// LS Electric XG5000 project: eduPJT_A
// PLC LSPLC
// module base 0 slot 0: 입출력 모듈:XBC-DR32H (DC 24V 입력, 릴레이 출력 32점)
// module base 0 slot 1: 입력 모듈:XBE-DC16A/B (DC24V 입력, 16점 / DC12/24V 입력, 16점)
// module base 0 slot 2: FEnet:XBL-EMTA (Ethernet 통신 모듈, 전기 Master)

PROGRAM 00_Global_Layer (task: 스캔 프로그램)

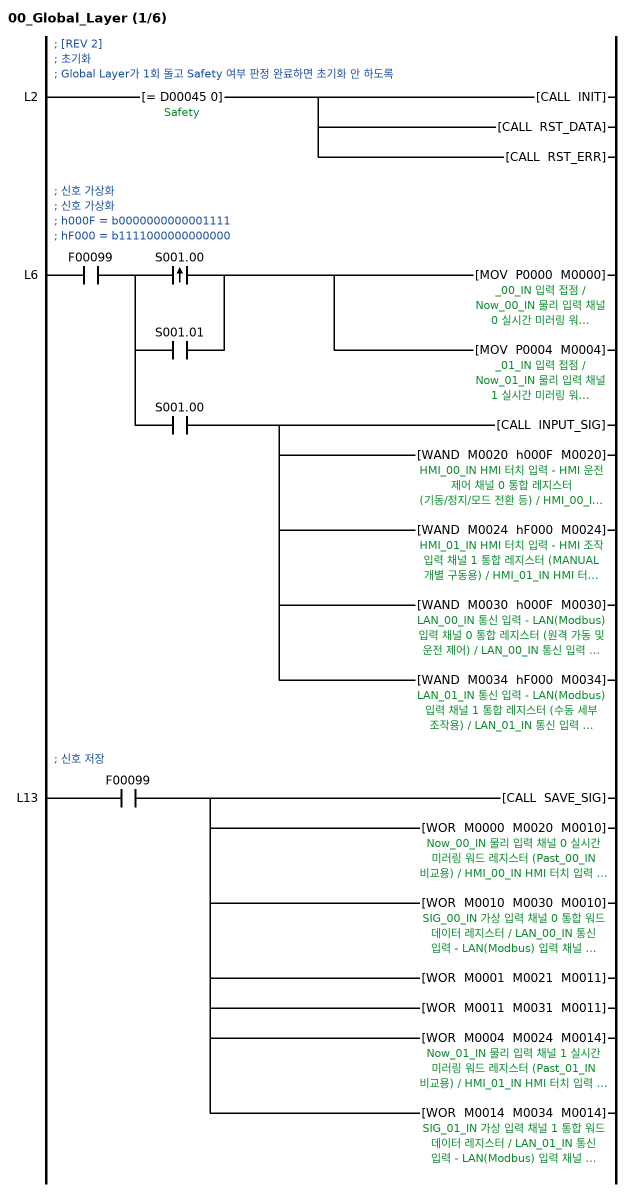
// [REV 2]
// 초기화
; L2
LOAD=     D00045 0	// Safety
CALL      INIT
CALL      RST_DATA
CALL      RST_ERR
// output comment: Global Layer가 1회 돌고 Safety 여부 판정 완료하면 초기화 안 하도록
// 신호 가상화
; L6
LOAD      F00099
MPUSH
LOADP     S001.00
OR        S001.01
AND LOAD
MOV       P0000 M0000	// _00_IN 입력 접점 / Now_00_IN 물리 입력 채널 0 실시간 미러링 워드 레지스터 (Past_00_IN 비교용)
MOV       P0004 M0004	// _01_IN 입력 접점 / Now_01_IN 물리 입력 채널 1 실시간 미러링 워드 레지스터 (Past_01_IN 비교용)
MPOP
AND       S001.00
CALL      INPUT_SIG
WAND      M0020 h000F M0020	// HMI_00_IN HMI 터치 입력 - HMI 운전 제어 채널 0 통합 레지스터 (기동/정지/모드 전환 등) / HMI_00_IN HMI 터치 입력 - HMI 운전 제어 채널 0 통합 레지스터 (기동/정지/모드 전환 등)
WAND      M0024 hF000 M0024	// HMI_01_IN HMI 터치 입력 - HMI 조작 입력 채널 1 통합 레지스터 (MANUAL 개별 구동용) / HMI_01_IN HMI 터치 입력 - HMI 조작 입력 채널 1 통합 레지스터 (MANUAL 개별 구동용)
WAND      M0030 h000F M0030	// LAN_00_IN 통신 입력 - LAN(Modbus) 입력 채널 0 통합 레지스터 (원격 가동 및 운전 제어) / LAN_00_IN 통신 입력 - LAN(Modbus) 입력 채널 0 통합 레지스터 (원격 가동 및 운전 제어)
WAND      M0034 hF000 M0034	// LAN_01_IN 통신 입력 - LAN(Modbus) 입력 채널 1 통합 레지스터 (수동 세부 조작용) / LAN_01_IN 통신 입력 - LAN(Modbus) 입력 채널 1 통합 레지스터 (수동 세부 조작용)
// output comment: 신호 가상화
// output comment: h000F = b0000000000001111
// output comment: hF000 = b1111000000000000
; L13
LOAD      F00099
CALL      SAVE_SIG
WOR       M0000 M0020 M0010	// Now_00_IN 물리 입력 채널 0 실시간 미러링 워드 레지스터 (Past_00_IN 비교용) / HMI_00_IN HMI 터치 입력 - HMI 운전 제어 채널 0 통합 레지스터 (기동/정지/모드 전환 등) / SIG_00_IN 가상 입력 채널 0 통합 워드 데이터 레지스터
WOR       M0010 M0030 M0010	// SIG_00_IN 가상 입력 채널 0 통합 워드 데이터 레지스터 / LAN_00_IN 통신 입력 - LAN(Modbus) 입력 채널 0 통합 레지스터 (원격 가동 및 운전 제어) / SIG_00_IN 가상 입력 채널 0 통합 워드 데이터 레지스터
WOR       M0001 M0021 M0011
WOR       M0011 M0031 M0011
WOR       M0004 M0024 M0014	// Now_01_IN 물리 입력 채널 1 실시간 미러링 워드 레지스터 (Past_01_IN 비교용) / HMI_01_IN HMI 터치 입력 - HMI 조작 입력 채널 1 통합 레지스터 (MANUAL 개별 구동용) / SIG_01_IN 가상 입력 채널 1 통합 워드 데이터 레지스터
WOR       M0014 M0034 M0014	// SIG_01_IN 가상 입력 채널 1 통합 워드 데이터 레지스터 / LAN_01_IN 통신 입력 - LAN(Modbus) 입력 채널 1 통합 레지스터 (수동 세부 조작용) / SIG_01_IN 가상 입력 채널 1 통합 워드 데이터 레지스터
// output comment: 신호 저장

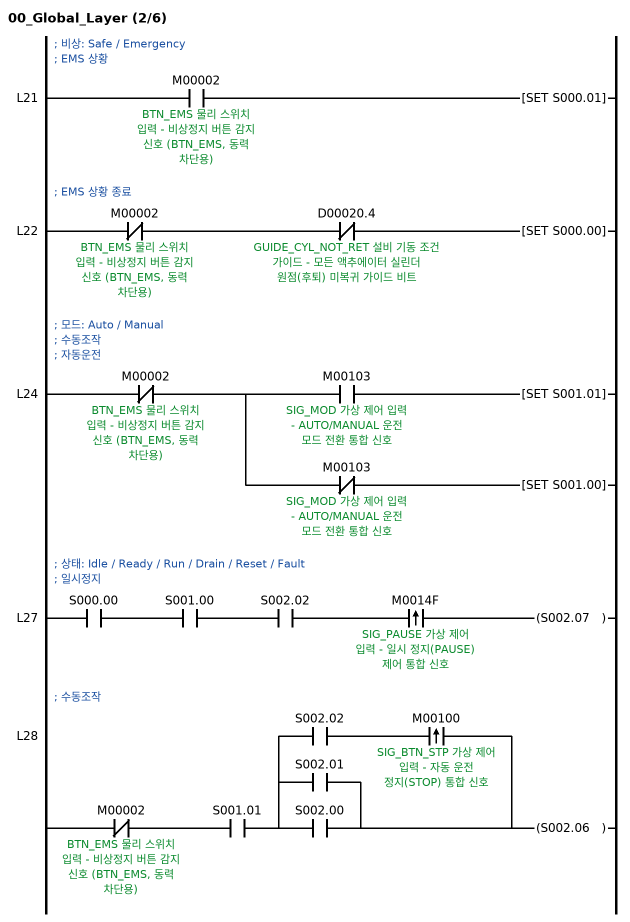
// 비상: Safe / Emergency
; L21
LOAD      M00002	// BTN_EMS 물리 스위치 입력 - 비상정지 버튼 감지 신호 (BTN_EMS, 동력 차단용)
SET       S000.01
// output comment: EMS 상황
; L22
LOAD NOT  M00002	// BTN_EMS 물리 스위치 입력 - 비상정지 버튼 감지 신호 (BTN_EMS, 동력 차단용)
AND NOT   D00020.4	// GUIDE_CYL_NOT_RET 설비 기동 조건 가이드 - 모든 액추에이터 실린더 원점(후퇴) 미복귀 가이드 비트
SET       S000.00
// output comment: EMS 상황 종료
// 모드: Auto / Manual
; L24
LOAD NOT  M00002	// BTN_EMS 물리 스위치 입력 - 비상정지 버튼 감지 신호 (BTN_EMS, 동력 차단용)
MPUSH
AND       M00103	// SIG_MOD 가상 제어 입력 - AUTO/MANUAL 운전 모드 전환 통합 신호
SET       S001.01
MPOP
AND NOT   M00103	// SIG_MOD 가상 제어 입력 - AUTO/MANUAL 운전 모드 전환 통합 신호
SET       S001.00
// output comment: 수동조작
// output comment: 자동운전
// 상태: Idle / Ready / Run / Drain / Reset / Fault
; L27
LOAD      S000.00
AND       S001.00
AND       S002.02
ANDP      M0014F	// SIG_PAUSE 가상 제어 입력 - 일시 정지(PAUSE) 제어 통합 신호
OUT       S002.07
// output comment: 일시정지
; L28
LOAD NOT  M00002	// BTN_EMS 물리 스위치 입력 - 비상정지 버튼 감지 신호 (BTN_EMS, 동력 차단용)
AND       S001.01
LOAD      S002.02
ANDP      M00100	// SIG_BTN_STP 가상 제어 입력 - 자동 운전 정지(STOP) 통합 신호
OR        S002.01
OR        S002.00
AND LOAD
OUT       S002.06
// output comment: 수동조작

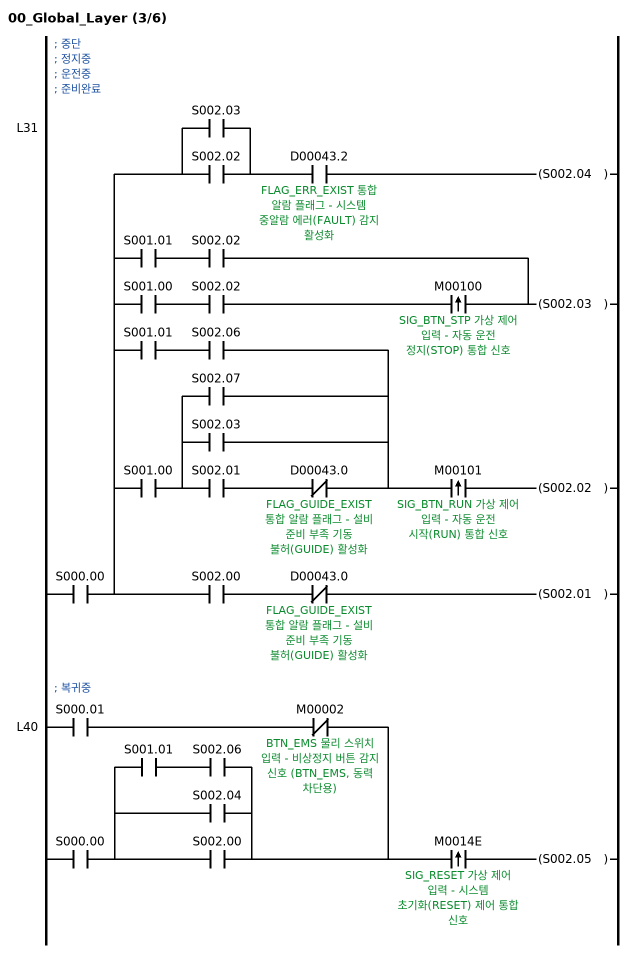
; L31
LOAD      S000.00
MPUSH
LOAD      S002.03
OR        S002.02
AND LOAD
AND       D00043.2	// FLAG_ERR_EXIST 통합 알람 플래그 - 시스템 중알람 에러(FAULT) 감지 활성화
OUT       S002.04
MLOAD
LOAD      S001.01
AND       S002.02
LOAD      S001.00
AND       S002.02
ANDP      M00100	// SIG_BTN_STP 가상 제어 입력 - 자동 운전 정지(STOP) 통합 신호
OR LOAD
AND LOAD
OUT       S002.03
MLOAD
LOAD      S001.01
AND       S002.06
LOAD      S001.00
LOAD      S002.07
OR        S002.03
LOAD      S002.01
AND NOT   D00043.0	// FLAG_GUIDE_EXIST 통합 알람 플래그 - 설비 준비 부족 기동 불허(GUIDE) 활성화
OR LOAD
AND LOAD
OR LOAD
AND LOAD
ANDP      M00101	// SIG_BTN_RUN 가상 제어 입력 - 자동 운전 시작(RUN) 통합 신호
OUT       S002.02
MPOP
AND       S002.00
AND NOT   D00043.0	// FLAG_GUIDE_EXIST 통합 알람 플래그 - 설비 준비 부족 기동 불허(GUIDE) 활성화
OUT       S002.01
// output comment: 중단
// output comment: 정지중
// output comment: 운전중
// output comment: 준비완료
; L40
LOAD      S000.01
AND NOT   M00002	// BTN_EMS 물리 스위치 입력 - 비상정지 버튼 감지 신호 (BTN_EMS, 동력 차단용)
LOAD      S000.00
LOAD      S001.01
AND       S002.06
OR        S002.04
OR        S002.00
AND LOAD
OR LOAD
ANDP      M0014E	// SIG_RESET 가상 제어 입력 - 시스템 초기화(RESET) 제어 통합 신호
OUT       S002.05
// output comment: 복귀중

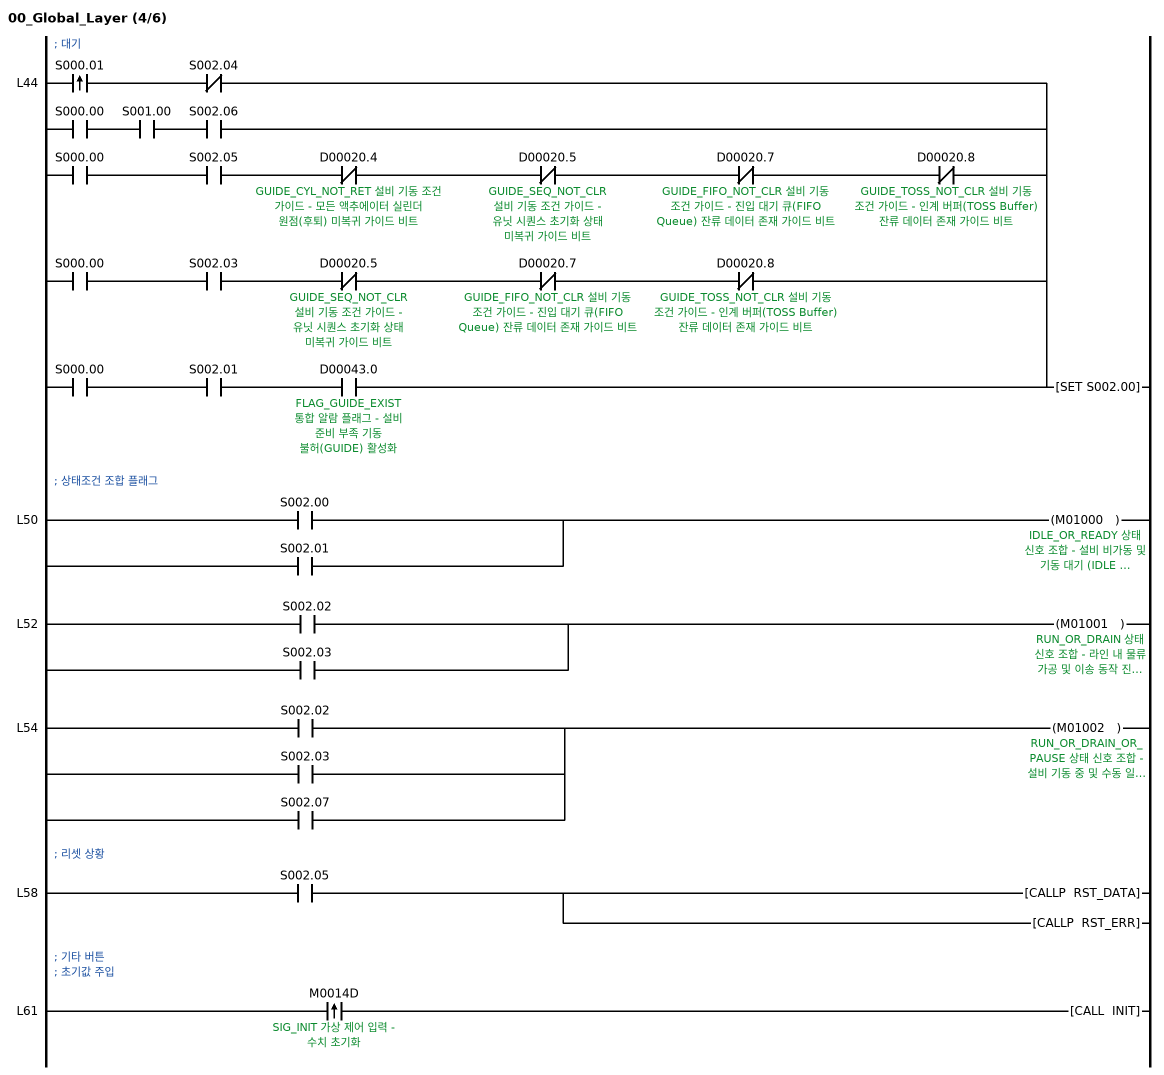
; L44
LOADP     S000.01
AND NOT   S002.04
LOAD      S000.00
AND       S001.00
AND       S002.06
OR LOAD
LOAD      S000.00
AND       S002.05
AND NOT   D00020.4	// GUIDE_CYL_NOT_RET 설비 기동 조건 가이드 - 모든 액추에이터 실린더 원점(후퇴) 미복귀 가이드 비트
AND NOT   D00020.5	// GUIDE_SEQ_NOT_CLR 설비 기동 조건 가이드 - 유닛 시퀀스 초기화 상태 미복귀 가이드 비트
AND NOT   D00020.7	// GUIDE_FIFO_NOT_CLR 설비 기동 조건 가이드 - 진입 대기 큐(FIFO Queue) 잔류 데이터 존재 가이드 비트
AND NOT   D00020.8	// GUIDE_TOSS_NOT_CLR 설비 기동 조건 가이드 - 인계 버퍼(TOSS Buffer) 잔류 데이터 존재 가이드 비트
OR LOAD
LOAD      S000.00
AND       S002.03
AND NOT   D00020.5	// GUIDE_SEQ_NOT_CLR 설비 기동 조건 가이드 - 유닛 시퀀스 초기화 상태 미복귀 가이드 비트
AND NOT   D00020.7	// GUIDE_FIFO_NOT_CLR 설비 기동 조건 가이드 - 진입 대기 큐(FIFO Queue) 잔류 데이터 존재 가이드 비트
AND NOT   D00020.8	// GUIDE_TOSS_NOT_CLR 설비 기동 조건 가이드 - 인계 버퍼(TOSS Buffer) 잔류 데이터 존재 가이드 비트
OR LOAD
LOAD      S000.00
AND       S002.01
AND       D00043.0	// FLAG_GUIDE_EXIST 통합 알람 플래그 - 설비 준비 부족 기동 불허(GUIDE) 활성화
OR LOAD
SET       S002.00
// output comment: 대기
// 상태조건 조합 플래그
; L50
LOAD      S002.00
OR        S002.01
OUT       M01000	// IDLE_OR_READY 상태 신호 조합 - 설비 비가동 및 기동 대기 (IDLE | READY) 플래그
; L52
LOAD      S002.02
OR        S002.03
OUT       M01001	// RUN_OR_DRAIN 상태 신호 조합 - 라인 내 물류 가공 및 이송 동작 진행 (RUN | DRAIN) 플래그
; L54
LOAD      S002.02
OR        S002.03
OR        S002.07
OUT       M01002	// RUN_OR_DRAIN_OR_PAUSE 상태 신호 조합 - 설비 기동 중 및 수동 일시 정지 (RUN | DRAIN | PAUSE) 플래그
// 리셋 상황
; L58
LOAD      S002.05
CALLP     RST_DATA
CALLP     RST_ERR
// 기타 버튼
; L61
LOADP     M0014D	// SIG_INIT 가상 제어 입력 - 수치 초기화
CALL      INIT
// output comment: 초기값 주입

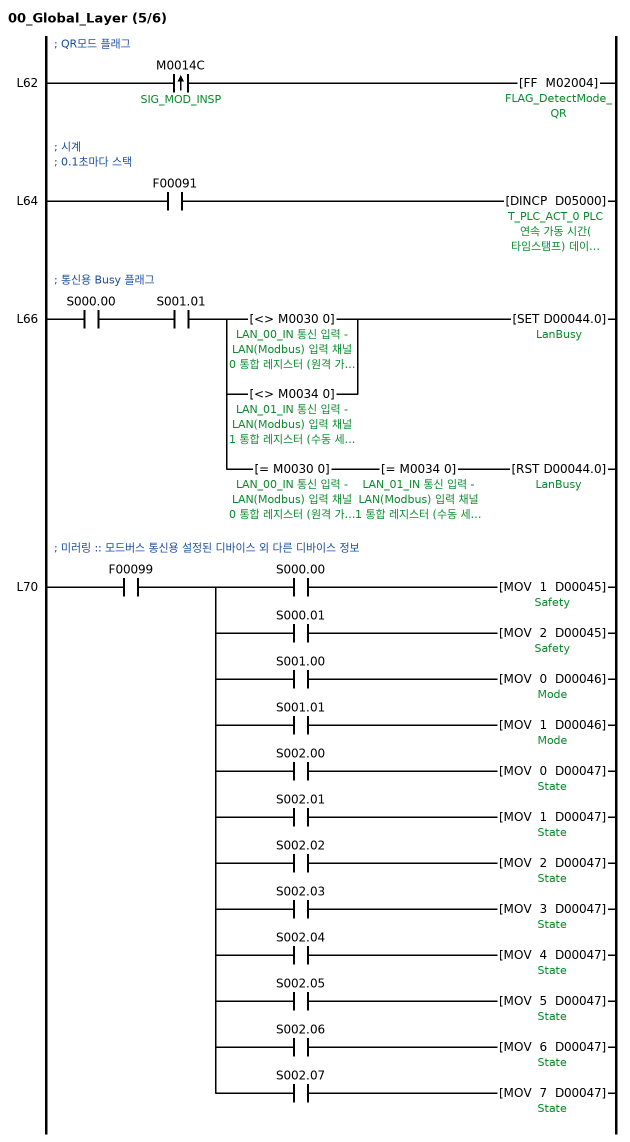
; L62
LOADP     M0014C	// SIG_MOD_INSP
FF        M02004	// FLAG_DetectMode_QR
// output comment: QR모드 플래그
// 시계
; L64
LOAD      F00091
DINCP     D05000	// T_PLC_ACT_0 PLC 연속 가동 시간(타임스탬프) 데이터 레지스터 하위 16비트 (0.1초 해상도)
// output comment: 0.1초마다 스택
// 통신용 Busy 플래그
; L66
LOAD      S000.00
AND       S001.01
MPUSH
LOAD<>    M0030 0	// LAN_00_IN 통신 입력 - LAN(Modbus) 입력 채널 0 통합 레지스터 (원격 가동 및 운전 제어)
OR<>      M0034 0	// LAN_01_IN 통신 입력 - LAN(Modbus) 입력 채널 1 통합 레지스터 (수동 세부 조작용)
AND LOAD
SET       D00044.0	// LanBusy
MPOP
AND=      M0030 0	// LAN_00_IN 통신 입력 - LAN(Modbus) 입력 채널 0 통합 레지스터 (원격 가동 및 운전 제어)
AND=      M0034 0	// LAN_01_IN 통신 입력 - LAN(Modbus) 입력 채널 1 통합 레지스터 (수동 세부 조작용)
RST       D00044.0	// LanBusy
// 미러링 :: 모드버스 통신용 설정된 디바이스 외 다른 디바이스 정보
; L70
LOAD      F00099
MPUSH
AND       S000.00
MOV       1 D00045	// Safety
MLOAD
AND       S000.01
MOV       2 D00045	// Safety
MLOAD
AND       S001.00
MOV       0 D00046	// Mode
MLOAD
AND       S001.01
MOV       1 D00046	// Mode
MLOAD
AND       S002.00
MOV       0 D00047	// State
MLOAD
AND       S002.01
MOV       1 D00047	// State
MLOAD
AND       S002.02
MOV       2 D00047	// State
MLOAD
AND       S002.03
MOV       3 D00047	// State
MLOAD
AND       S002.04
MOV       4 D00047	// State
MLOAD
AND       S002.05
MOV       5 D00047	// State
MLOAD
AND       S002.06
MOV       6 D00047	// State
MPOP
AND       S002.07
MOV       7 D00047	// State

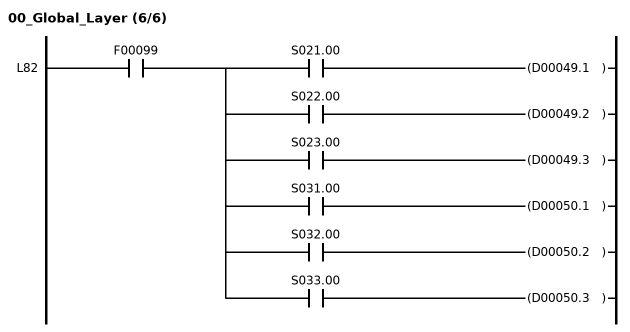
; L82
LOAD      F00099
MPUSH
AND       S021.00
OUT       D00049.1
MLOAD
AND       S022.00
OUT       D00049.2
MLOAD
AND       S023.00
OUT       D00049.3
MLOAD
AND       S031.00
OUT       D00050.1
MLOAD
AND       S032.00
OUT       D00050.2
MPOP
AND       S033.00
OUT       D00050.3

PROGRAM 01_Sequence_Layer (task: 스캔 프로그램)

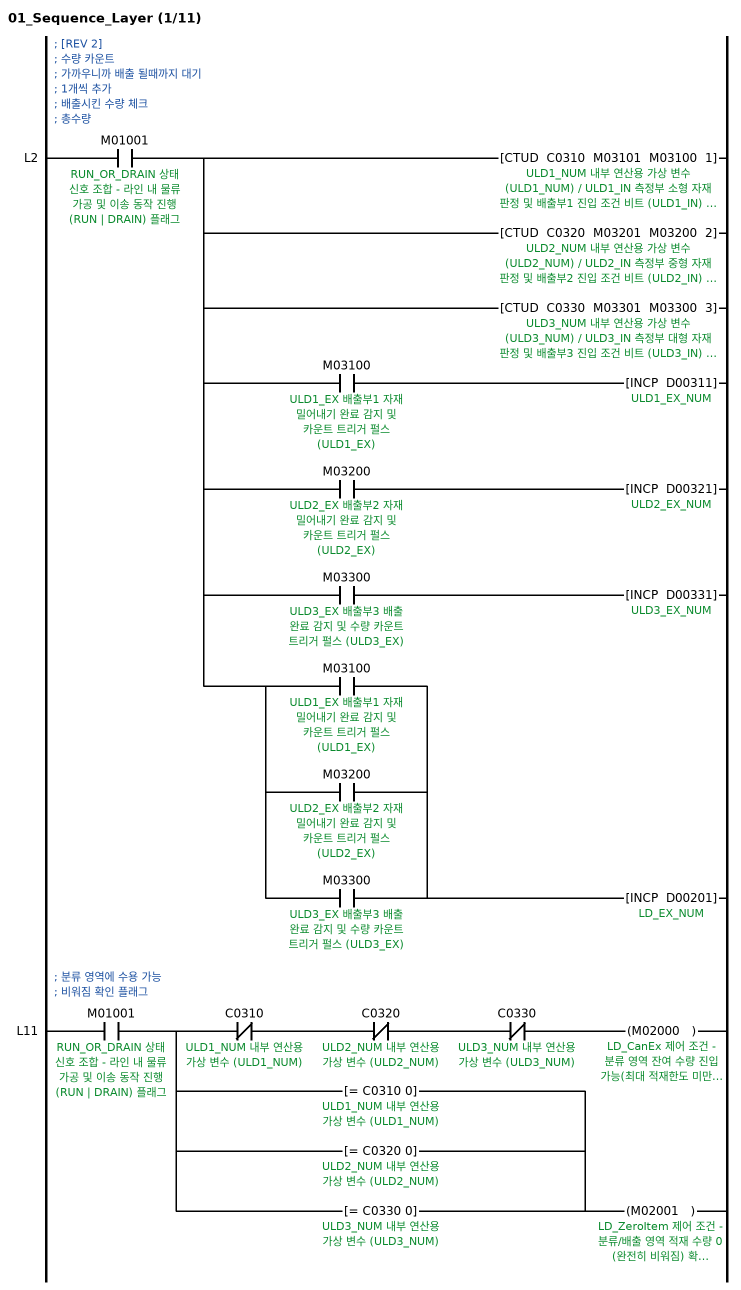
// [REV 2]
// 수량 카운트
; L2
LOAD      M01001	// RUN_OR_DRAIN 상태 신호 조합 - 라인 내 물류 가공 및 이송 동작 진행 (RUN | DRAIN) 플래그
CTUD      C0310 M03101 M03100 1	// ULD1_NUM 내부 연산용 가상 변수 (ULD1_NUM) / ULD1_IN 측정부 소형 자재 판정 및 배출부1 진입 조건 비트 (ULD1_IN) / ULD1_EX 배출부1 자재 밀어내기 완료 감지 및 카운트 트리거 펄스 (ULD1_EX)
CTUD      C0320 M03201 M03200 2	// ULD2_NUM 내부 연산용 가상 변수 (ULD2_NUM) / ULD2_IN 측정부 중형 자재 판정 및 배출부2 진입 조건 비트 (ULD2_IN) / ULD2_EX 배출부2 자재 밀어내기 완료 감지 및 카운트 트리거 펄스 (ULD2_EX)
CTUD      C0330 M03301 M03300 3	// ULD3_NUM 내부 연산용 가상 변수 (ULD3_NUM) / ULD3_IN 측정부 대형 자재 판정 및 배출부3 진입 조건 비트 (ULD3_IN) / ULD3_EX 배출부3 배출 완료 감지 및 수량 카운트 트리거 펄스 (ULD3_EX)
MPUSH
AND       M03100	// ULD1_EX 배출부1 자재 밀어내기 완료 감지 및 카운트 트리거 펄스 (ULD1_EX)
INCP      D00311	// ULD1_EX_NUM
MLOAD
AND       M03200	// ULD2_EX 배출부2 자재 밀어내기 완료 감지 및 카운트 트리거 펄스 (ULD2_EX)
INCP      D00321	// ULD2_EX_NUM
MLOAD
AND       M03300	// ULD3_EX 배출부3 배출 완료 감지 및 수량 카운트 트리거 펄스 (ULD3_EX)
INCP      D00331	// ULD3_EX_NUM
MPOP
LOAD      M03100	// ULD1_EX 배출부1 자재 밀어내기 완료 감지 및 카운트 트리거 펄스 (ULD1_EX)
OR        M03200	// ULD2_EX 배출부2 자재 밀어내기 완료 감지 및 카운트 트리거 펄스 (ULD2_EX)
OR        M03300	// ULD3_EX 배출부3 배출 완료 감지 및 수량 카운트 트리거 펄스 (ULD3_EX)
AND LOAD
INCP      D00201	// LD_EX_NUM
// output comment: 가까우니까 배출 될때까지 대기
// output comment: 1개씩 추가
// output comment: 배출시킨 수량 체크
// output comment: 총수량
; L11
LOAD      M01001	// RUN_OR_DRAIN 상태 신호 조합 - 라인 내 물류 가공 및 이송 동작 진행 (RUN | DRAIN) 플래그
MPUSH
AND NOT   C0310	// ULD1_NUM 내부 연산용 가상 변수 (ULD1_NUM)
AND NOT   C0320	// ULD2_NUM 내부 연산용 가상 변수 (ULD2_NUM)
AND NOT   C0330	// ULD3_NUM 내부 연산용 가상 변수 (ULD3_NUM)
OUT       M02000	// LD_CanEx 제어 조건 - 분류 영역 잔여 수량 진입 가능(최대 적재한도 미만) 확인 플래그 (LD_CanEx)
MPOP
LOAD=     C0310 0	// ULD1_NUM 내부 연산용 가상 변수 (ULD1_NUM)
OR=       C0320 0	// ULD2_NUM 내부 연산용 가상 변수 (ULD2_NUM)
OR=       C0330 0	// ULD3_NUM 내부 연산용 가상 변수 (ULD3_NUM)
AND LOAD
OUT       M02001	// LD_ZeroItem 제어 조건 - 분류/배출 영역 적재 수량 0 (완전히 비워짐) 확인 플래그 (LD_ZeroItem)
// output comment: 분류 영역에 수용 가능
// output comment: 비워짐 확인 플래그

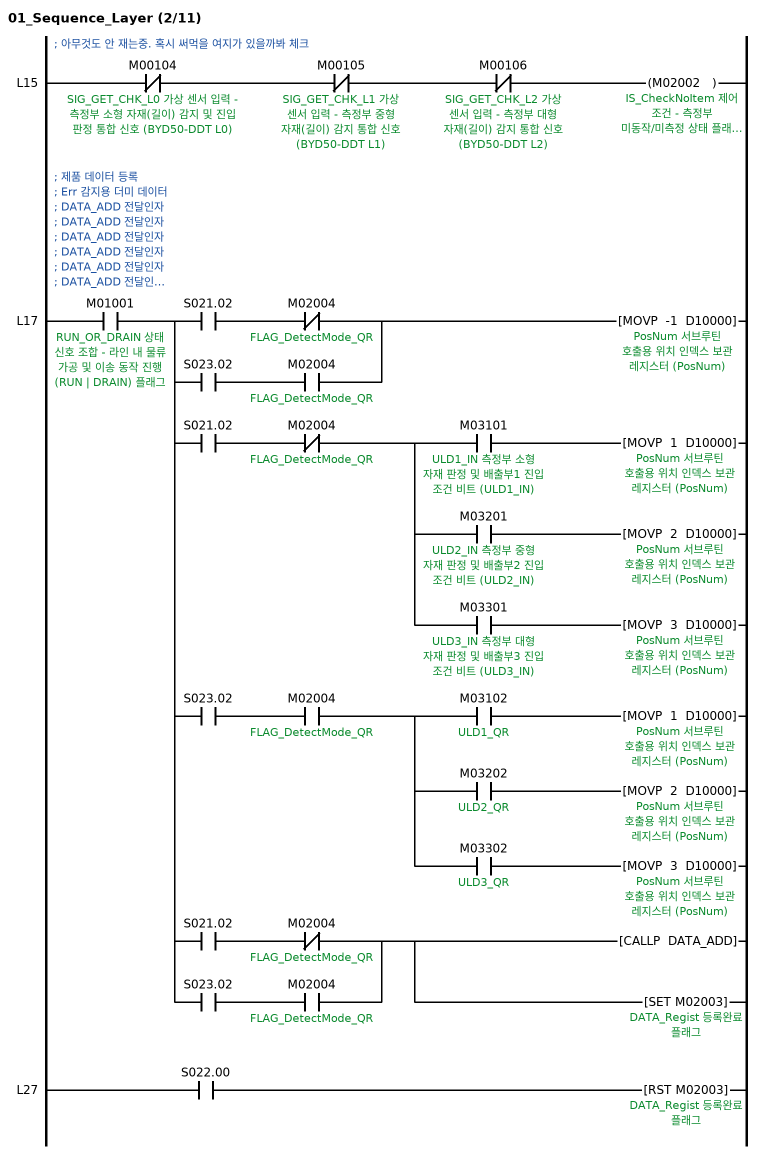
; L15
LOAD NOT  M00104	// SIG_GET_CHK_L0 가상 센서 입력 - 측정부 소형 자재(길이) 감지 및 진입 판정 통합 신호 (BYD50-DDT L0)
AND NOT   M00105	// SIG_GET_CHK_L1 가상 센서 입력 - 측정부 중형 자재(길이) 감지 통합 신호 (BYD50-DDT L1)
AND NOT   M00106	// SIG_GET_CHK_L2 가상 센서 입력 - 측정부 대형 자재(길이) 감지 통합 신호 (BYD50-DDT L2)
OUT       M02002	// IS_CheckNoItem 제어 조건 - 측정부 미동작/미측정 상태 플래그 (IS_CheckNoItem)
// output comment: 아무것도 안 재는중. 혹시 써먹을 여지가 있을까봐 체크
// 제품 데이터 등록
; L17
LOAD      M01001	// RUN_OR_DRAIN 상태 신호 조합 - 라인 내 물류 가공 및 이송 동작 진행 (RUN | DRAIN) 플래그
MPUSH
LOAD      S021.02
AND NOT   M02004	// FLAG_DetectMode_QR
LOAD      S023.02
AND       M02004	// FLAG_DetectMode_QR
OR LOAD
AND LOAD
MOVP      -1 D10000	// PosNum 서브루틴 호출용 위치 인덱스 보관 레지스터 (PosNum)
MLOAD
AND       S021.02
AND NOT   M02004	// FLAG_DetectMode_QR
MPUSH
AND       M03101	// ULD1_IN 측정부 소형 자재 판정 및 배출부1 진입 조건 비트 (ULD1_IN)
MOVP      1 D10000	// PosNum 서브루틴 호출용 위치 인덱스 보관 레지스터 (PosNum)
MLOAD
AND       M03201	// ULD2_IN 측정부 중형 자재 판정 및 배출부2 진입 조건 비트 (ULD2_IN)
MOVP      2 D10000	// PosNum 서브루틴 호출용 위치 인덱스 보관 레지스터 (PosNum)
MPOP
AND       M03301	// ULD3_IN 측정부 대형 자재 판정 및 배출부3 진입 조건 비트 (ULD3_IN)
MOVP      3 D10000	// PosNum 서브루틴 호출용 위치 인덱스 보관 레지스터 (PosNum)
MLOAD
AND       S023.02
AND       M02004	// FLAG_DetectMode_QR
MPUSH
AND       M03102	// ULD1_QR
MOVP      1 D10000	// PosNum 서브루틴 호출용 위치 인덱스 보관 레지스터 (PosNum)
MLOAD
AND       M03202	// ULD2_QR
MOVP      2 D10000	// PosNum 서브루틴 호출용 위치 인덱스 보관 레지스터 (PosNum)
MPOP
AND       M03302	// ULD3_QR
MOVP      3 D10000	// PosNum 서브루틴 호출용 위치 인덱스 보관 레지스터 (PosNum)
MPOP
LOAD      S021.02
AND NOT   M02004	// FLAG_DetectMode_QR
LOAD      S023.02
AND       M02004	// FLAG_DetectMode_QR
OR LOAD
AND LOAD
CALLP     DATA_ADD
SET       M02003	// DATA_Regist 등록완료 플래그
// output comment: Err 감지용 더미 데이터
// output comment: DATA_ADD 전달인자
// output comment: DATA_ADD 전달인자
// output comment: DATA_ADD 전달인자
// output comment: DATA_ADD 전달인자
// output comment: DATA_ADD 전달인자
// output comment: DATA_ADD 전달인자
// output comment: 선입선출 데이터 입력
// output comment: 등록완료 플래그
; L27
LOAD      S022.00
RST       M02003	// DATA_Regist 등록완료 플래그

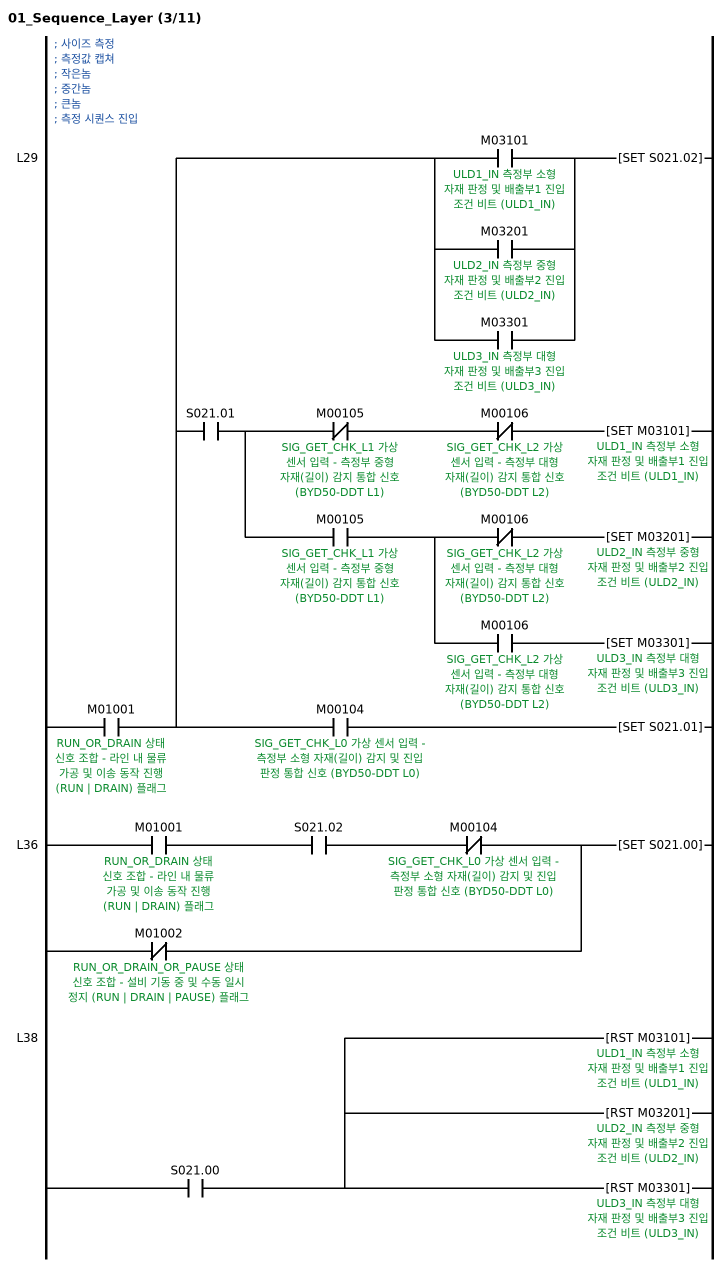
// 
// 사이즈 측정
; L29
LOAD      M01001	// RUN_OR_DRAIN 상태 신호 조합 - 라인 내 물류 가공 및 이송 동작 진행 (RUN | DRAIN) 플래그
MPUSH
LOAD      M03101	// ULD1_IN 측정부 소형 자재 판정 및 배출부1 진입 조건 비트 (ULD1_IN)
OR        M03201	// ULD2_IN 측정부 중형 자재 판정 및 배출부2 진입 조건 비트 (ULD2_IN)
OR        M03301	// ULD3_IN 측정부 대형 자재 판정 및 배출부3 진입 조건 비트 (ULD3_IN)
AND LOAD
SET       S021.02
MLOAD
AND       S021.01
MPUSH
AND NOT   M00105	// SIG_GET_CHK_L1 가상 센서 입력 - 측정부 중형 자재(길이) 감지 통합 신호 (BYD50-DDT L1)
AND NOT   M00106	// SIG_GET_CHK_L2 가상 센서 입력 - 측정부 대형 자재(길이) 감지 통합 신호 (BYD50-DDT L2)
SET       M03101	// ULD1_IN 측정부 소형 자재 판정 및 배출부1 진입 조건 비트 (ULD1_IN)
MPOP
AND       M00105	// SIG_GET_CHK_L1 가상 센서 입력 - 측정부 중형 자재(길이) 감지 통합 신호 (BYD50-DDT L1)
MPUSH
AND NOT   M00106	// SIG_GET_CHK_L2 가상 센서 입력 - 측정부 대형 자재(길이) 감지 통합 신호 (BYD50-DDT L2)
SET       M03201	// ULD2_IN 측정부 중형 자재 판정 및 배출부2 진입 조건 비트 (ULD2_IN)
MPOP
AND       M00106	// SIG_GET_CHK_L2 가상 센서 입력 - 측정부 대형 자재(길이) 감지 통합 신호 (BYD50-DDT L2)
SET       M03301	// ULD3_IN 측정부 대형 자재 판정 및 배출부3 진입 조건 비트 (ULD3_IN)
MPOP
AND       M00104	// SIG_GET_CHK_L0 가상 센서 입력 - 측정부 소형 자재(길이) 감지 및 진입 판정 통합 신호 (BYD50-DDT L0)
SET       S021.01
// output comment: 측정값 캡쳐
// output comment: 작은놈
// output comment: 중간놈
// output comment: 큰놈
// output comment: 측정 시퀀스 진입
; L36
LOAD      M01001	// RUN_OR_DRAIN 상태 신호 조합 - 라인 내 물류 가공 및 이송 동작 진행 (RUN | DRAIN) 플래그
AND       S021.02
AND NOT   M00104	// SIG_GET_CHK_L0 가상 센서 입력 - 측정부 소형 자재(길이) 감지 및 진입 판정 통합 신호 (BYD50-DDT L0)
OR NOT    M01002	// RUN_OR_DRAIN_OR_PAUSE 상태 신호 조합 - 설비 기동 중 및 수동 일시 정지 (RUN | DRAIN | PAUSE) 플래그
SET       S021.00
; L38
LOAD      S021.00
RST       M03101	// ULD1_IN 측정부 소형 자재 판정 및 배출부1 진입 조건 비트 (ULD1_IN)
RST       M03201	// ULD2_IN 측정부 중형 자재 판정 및 배출부2 진입 조건 비트 (ULD2_IN)
RST       M03301	// ULD3_IN 측정부 대형 자재 판정 및 배출부3 진입 조건 비트 (ULD3_IN)

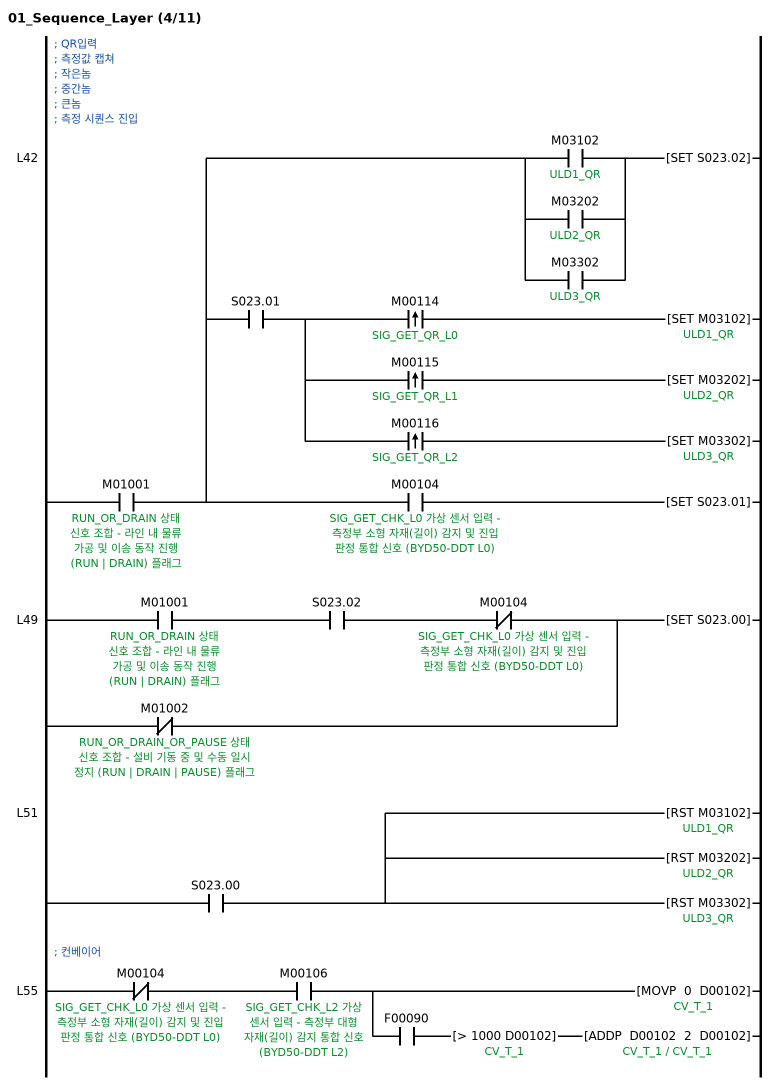
// QR입력
; L42
LOAD      M01001	// RUN_OR_DRAIN 상태 신호 조합 - 라인 내 물류 가공 및 이송 동작 진행 (RUN | DRAIN) 플래그
MPUSH
LOAD      M03102	// ULD1_QR
OR        M03202	// ULD2_QR
OR        M03302	// ULD3_QR
AND LOAD
SET       S023.02
MLOAD
AND       S023.01
MPUSH
ANDP      M00114	// SIG_GET_QR_L0
SET       M03102	// ULD1_QR
MLOAD
ANDP      M00115	// SIG_GET_QR_L1
SET       M03202	// ULD2_QR
MPOP
ANDP      M00116	// SIG_GET_QR_L2
SET       M03302	// ULD3_QR
MPOP
AND       M00104	// SIG_GET_CHK_L0 가상 센서 입력 - 측정부 소형 자재(길이) 감지 및 진입 판정 통합 신호 (BYD50-DDT L0)
SET       S023.01
// output comment: 측정값 캡쳐
// output comment: 작은놈
// output comment: 중간놈
// output comment: 큰놈
// output comment: 측정 시퀀스 진입
; L49
LOAD      M01001	// RUN_OR_DRAIN 상태 신호 조합 - 라인 내 물류 가공 및 이송 동작 진행 (RUN | DRAIN) 플래그
AND       S023.02
AND NOT   M00104	// SIG_GET_CHK_L0 가상 센서 입력 - 측정부 소형 자재(길이) 감지 및 진입 판정 통합 신호 (BYD50-DDT L0)
OR NOT    M01002	// RUN_OR_DRAIN_OR_PAUSE 상태 신호 조합 - 설비 기동 중 및 수동 일시 정지 (RUN | DRAIN | PAUSE) 플래그
SET       S023.00
; L51
LOAD      S023.00
RST       M03102	// ULD1_QR
RST       M03202	// ULD2_QR
RST       M03302	// ULD3_QR
// 
// 컨베이어
; L55
LOAD NOT  M00104	// SIG_GET_CHK_L0 가상 센서 입력 - 측정부 소형 자재(길이) 감지 및 진입 판정 통합 신호 (BYD50-DDT L0)
AND       M00106	// SIG_GET_CHK_L2 가상 센서 입력 - 측정부 대형 자재(길이) 감지 통합 신호 (BYD50-DDT L2)
MOVP      0 D00102	// CV_T_1
AND       F00090
AND>      1000 D00102	// CV_T_1
ADDP      D00102 2 D00102	// CV_T_1 / CV_T_1

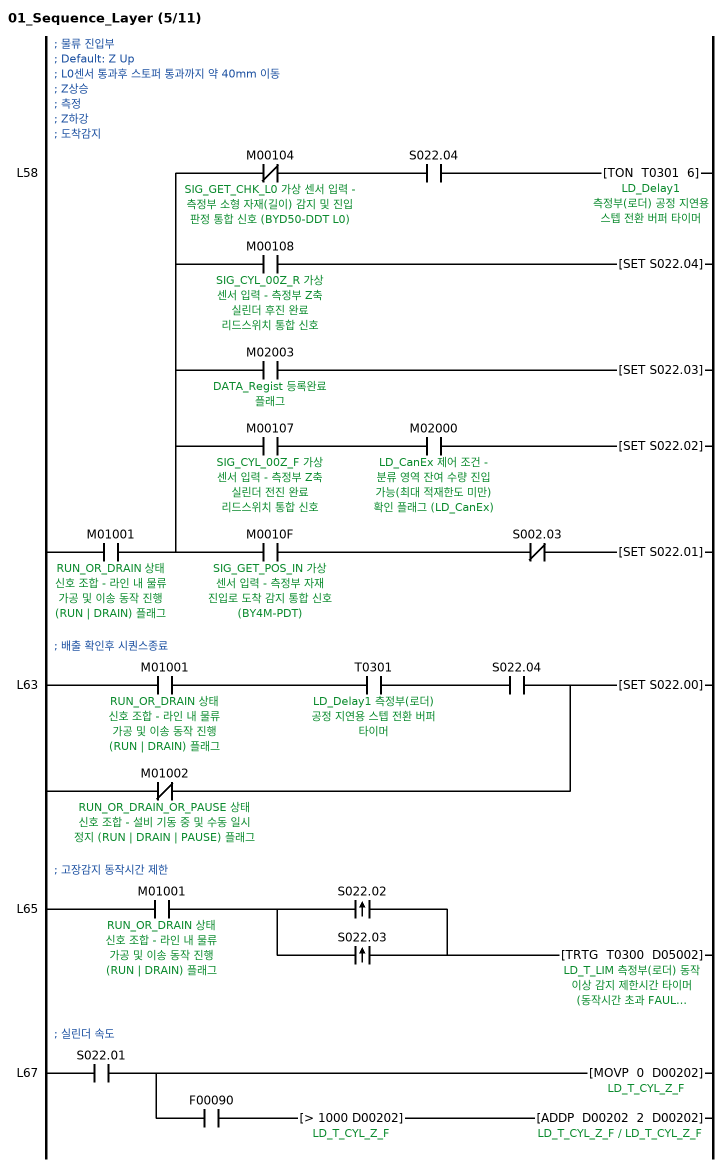
// 
// 물류 진입부
// 
// Default: Z Up
; L58
LOAD      M01001	// RUN_OR_DRAIN 상태 신호 조합 - 라인 내 물류 가공 및 이송 동작 진행 (RUN | DRAIN) 플래그
MPUSH
AND NOT   M00104	// SIG_GET_CHK_L0 가상 센서 입력 - 측정부 소형 자재(길이) 감지 및 진입 판정 통합 신호 (BYD50-DDT L0)
AND       S022.04
TON       T0301 6	// LD_Delay1 측정부(로더) 공정 지연용 스텝 전환 버퍼 타이머
MLOAD
AND       M00108	// SIG_CYL_00Z_R 가상 센서 입력 - 측정부 Z축 실린더 후진 완료 리드스위치 통합 신호
SET       S022.04
MLOAD
AND       M02003	// DATA_Regist 등록완료 플래그
SET       S022.03
MLOAD
AND       M00107	// SIG_CYL_00Z_F 가상 센서 입력 - 측정부 Z축 실린더 전진 완료 리드스위치 통합 신호
AND       M02000	// LD_CanEx 제어 조건 - 분류 영역 잔여 수량 진입 가능(최대 적재한도 미만) 확인 플래그 (LD_CanEx)
SET       S022.02
MPOP
AND       M0010F	// SIG_GET_POS_IN 가상 센서 입력 - 측정부 자재 진입로 도착 감지 통합 신호 (BY4M-PDT)
AND NOT   S002.03
SET       S022.01
// output comment: L0센서 통과후 스토퍼 통과까지 약 40mm 이동
// output comment: Z상승
// output comment: 측정
// output comment: Z하강
// output comment: 도착감지
; L63
LOAD      M01001	// RUN_OR_DRAIN 상태 신호 조합 - 라인 내 물류 가공 및 이송 동작 진행 (RUN | DRAIN) 플래그
AND       T0301	// LD_Delay1 측정부(로더) 공정 지연용 스텝 전환 버퍼 타이머
AND       S022.04
OR NOT    M01002	// RUN_OR_DRAIN_OR_PAUSE 상태 신호 조합 - 설비 기동 중 및 수동 일시 정지 (RUN | DRAIN | PAUSE) 플래그
SET       S022.00
// output comment: 배출 확인후 시퀀스종료
; L65
LOAD      M01001	// RUN_OR_DRAIN 상태 신호 조합 - 라인 내 물류 가공 및 이송 동작 진행 (RUN | DRAIN) 플래그
LOADP     S022.02
ORP       S022.03
AND LOAD
TRTG      T0300 D05002	// LD_T_LIM 측정부(로더) 동작 이상 감지 제한시간 타이머 (동작시간 초과 FAULT 트리거) / T_Limit 단위 동작 고장 감지 제한시간(타임아웃) 기준값 설정 레지스터
// output comment: 고장감지 동작시간 제한
; L67
LOAD      S022.01
MOVP      0 D00202	// LD_T_CYL_Z_F
AND       F00090
AND>      1000 D00202	// LD_T_CYL_Z_F
ADDP      D00202 2 D00202	// LD_T_CYL_Z_F / LD_T_CYL_Z_F
// output comment: 실린더 속도

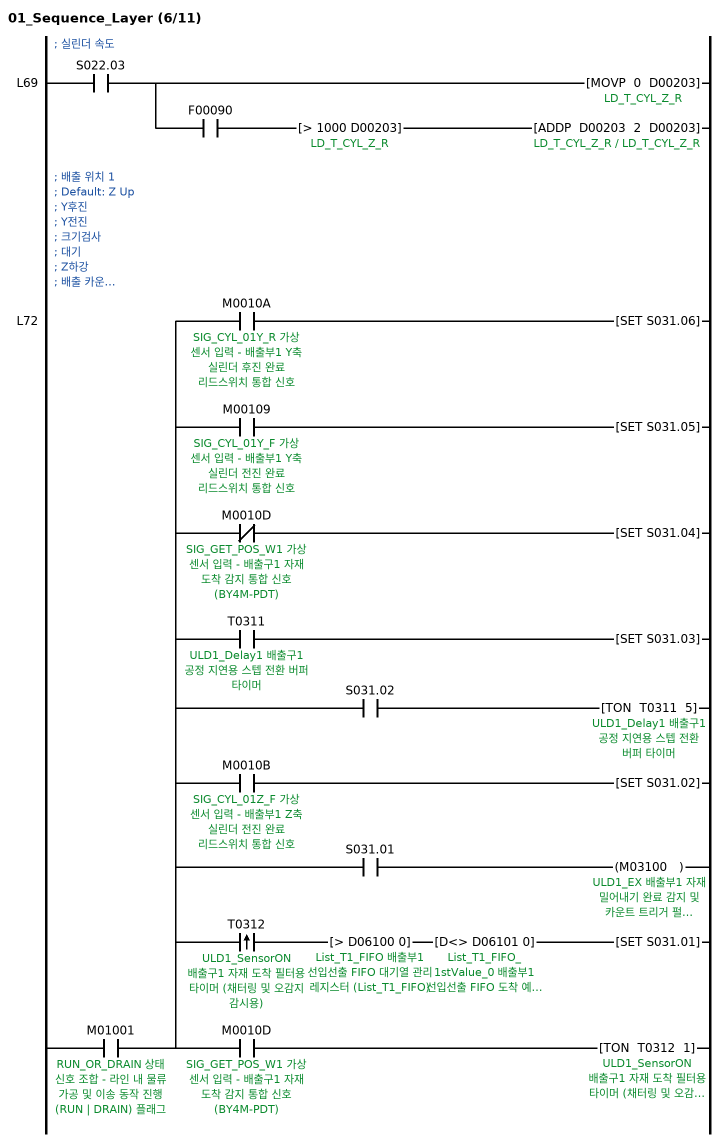
; L69
LOAD      S022.03
MOVP      0 D00203	// LD_T_CYL_Z_R
AND       F00090
AND>      1000 D00203	// LD_T_CYL_Z_R
ADDP      D00203 2 D00203	// LD_T_CYL_Z_R / LD_T_CYL_Z_R
// output comment: 실린더 속도
// 
// 배출 위치 1
// 
// Default: Z Up
; L72
LOAD      M01001	// RUN_OR_DRAIN 상태 신호 조합 - 라인 내 물류 가공 및 이송 동작 진행 (RUN | DRAIN) 플래그
MPUSH
AND       M0010A	// SIG_CYL_01Y_R 가상 센서 입력 - 배출부1 Y축 실린더 후진 완료 리드스위치 통합 신호
SET       S031.06
MLOAD
AND       M00109	// SIG_CYL_01Y_F 가상 센서 입력 - 배출부1 Y축 실린더 전진 완료 리드스위치 통합 신호
SET       S031.05
MLOAD
AND NOT   M0010D	// SIG_GET_POS_W1 가상 센서 입력 - 배출구1 자재 도착 감지 통합 신호 (BY4M-PDT)
SET       S031.04
MLOAD
AND       T0311	// ULD1_Delay1 배출구1 공정 지연용 스텝 전환 버퍼 타이머
SET       S031.03
MLOAD
AND       S031.02
TON       T0311 5	// ULD1_Delay1 배출구1 공정 지연용 스텝 전환 버퍼 타이머
MLOAD
AND       M0010B	// SIG_CYL_01Z_F 가상 센서 입력 - 배출부1 Z축 실린더 전진 완료 리드스위치 통합 신호
SET       S031.02
MLOAD
AND       S031.01
OUT       M03100	// ULD1_EX 배출부1 자재 밀어내기 완료 감지 및 카운트 트리거 펄스 (ULD1_EX)
MLOAD
ANDP      T0312	// ULD1_SensorON 배출구1 자재 도착 필터용 타이머 (채터링 및 오감지 감시용)
AND>      D06100 0	// List_T1_FIFO 배출부1 선입선출 FIFO 대기열 관리 레지스터 (List_T1_FIFO)
ANDD<>    D06101 0	// List_T1_FIFO_1stValue_0 배출부1 선입선출 FIFO 도착 예정 시간 데이터 레지스터 하위 16비트 (32비트 연산)
SET       S031.01
MPOP
AND       M0010D	// SIG_GET_POS_W1 가상 센서 입력 - 배출구1 자재 도착 감지 통합 신호 (BY4M-PDT)
TON       T0312 1	// ULD1_SensorON 배출구1 자재 도착 필터용 타이머 (채터링 및 오감지 감시용)
// output comment: Y후진
// output comment: Y전진
// output comment: 크기검사
// output comment: 대기
// output comment: Z하강
// output comment: 배출 카운트
// output comment: 도착감지
// output comment: 채터링->데이터오염 방지

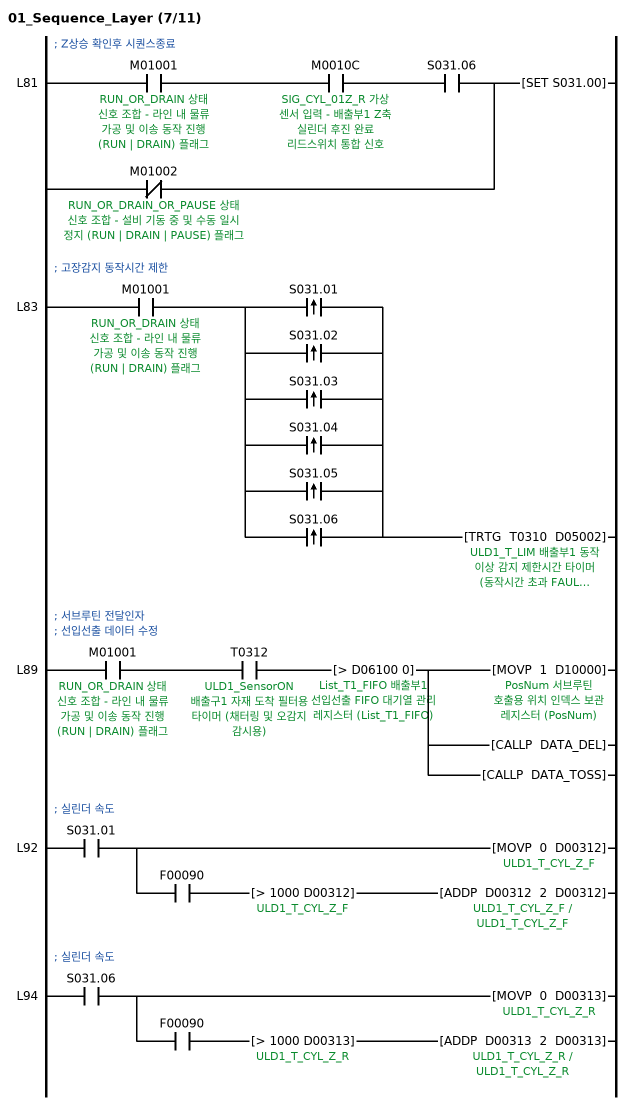
; L81
LOAD      M01001	// RUN_OR_DRAIN 상태 신호 조합 - 라인 내 물류 가공 및 이송 동작 진행 (RUN | DRAIN) 플래그
AND       M0010C	// SIG_CYL_01Z_R 가상 센서 입력 - 배출부1 Z축 실린더 후진 완료 리드스위치 통합 신호
AND       S031.06
OR NOT    M01002	// RUN_OR_DRAIN_OR_PAUSE 상태 신호 조합 - 설비 기동 중 및 수동 일시 정지 (RUN | DRAIN | PAUSE) 플래그
SET       S031.00
// output comment: Z상승 확인후 시퀀스종료
; L83
LOAD      M01001	// RUN_OR_DRAIN 상태 신호 조합 - 라인 내 물류 가공 및 이송 동작 진행 (RUN | DRAIN) 플래그
LOADP     S031.01
ORP       S031.02
ORP       S031.03
ORP       S031.04
ORP       S031.05
ORP       S031.06
AND LOAD
TRTG      T0310 D05002	// ULD1_T_LIM 배출부1 동작 이상 감지 제한시간 타이머 (동작시간 초과 FAULT 트리거) / T_Limit 단위 동작 고장 감지 제한시간(타임아웃) 기준값 설정 레지스터
// output comment: 고장감지 동작시간 제한
; L89
LOAD      M01001	// RUN_OR_DRAIN 상태 신호 조합 - 라인 내 물류 가공 및 이송 동작 진행 (RUN | DRAIN) 플래그
AND       T0312	// ULD1_SensorON 배출구1 자재 도착 필터용 타이머 (채터링 및 오감지 감시용)
AND>      D06100 0	// List_T1_FIFO 배출부1 선입선출 FIFO 대기열 관리 레지스터 (List_T1_FIFO)
MOVP      1 D10000	// PosNum 서브루틴 호출용 위치 인덱스 보관 레지스터 (PosNum)
CALLP     DATA_DEL
CALLP     DATA_TOSS
// output comment: 서브루틴 전달인자
// output comment: 선입선출 데이터 수정
; L92
LOAD      S031.01
MOVP      0 D00312	// ULD1_T_CYL_Z_F
AND       F00090
AND>      1000 D00312	// ULD1_T_CYL_Z_F
ADDP      D00312 2 D00312	// ULD1_T_CYL_Z_F / ULD1_T_CYL_Z_F
// output comment: 실린더 속도
; L94
LOAD      S031.06
MOVP      0 D00313	// ULD1_T_CYL_Z_R
AND       F00090
AND>      1000 D00313	// ULD1_T_CYL_Z_R
ADDP      D00313 2 D00313	// ULD1_T_CYL_Z_R / ULD1_T_CYL_Z_R
// output comment: 실린더 속도

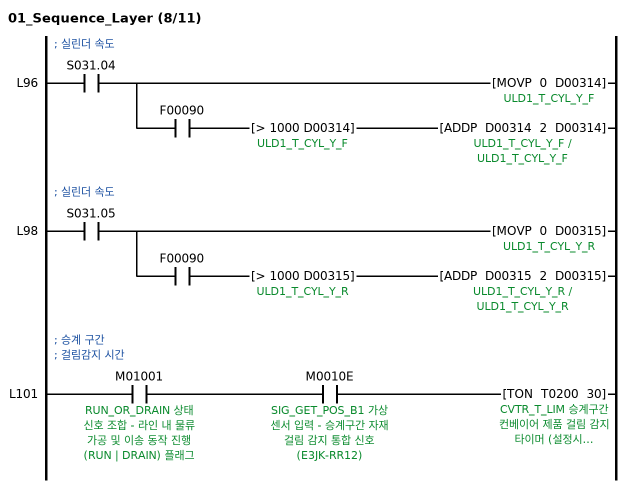
; L96
LOAD      S031.04
MOVP      0 D00314	// ULD1_T_CYL_Y_F
AND       F00090
AND>      1000 D00314	// ULD1_T_CYL_Y_F
ADDP      D00314 2 D00314	// ULD1_T_CYL_Y_F / ULD1_T_CYL_Y_F
// output comment: 실린더 속도
; L98
LOAD      S031.05
MOVP      0 D00315	// ULD1_T_CYL_Y_R
AND       F00090
AND>      1000 D00315	// ULD1_T_CYL_Y_R
ADDP      D00315 2 D00315	// ULD1_T_CYL_Y_R / ULD1_T_CYL_Y_R
// output comment: 실린더 속도
// 승계 구간
; L101
LOAD      M01001	// RUN_OR_DRAIN 상태 신호 조합 - 라인 내 물류 가공 및 이송 동작 진행 (RUN | DRAIN) 플래그
AND       M0010E	// SIG_GET_POS_B1 가상 센서 입력 - 승계구간 자재 걸림 감지 통합 신호 (E3JK-RR12)
TON       T0200 30	// CVTR_T_LIM 승계구간 컨베이어 제품 걸림 감지 타이머 (설정시간 30.0초)
// output comment: 걸림감지 시간

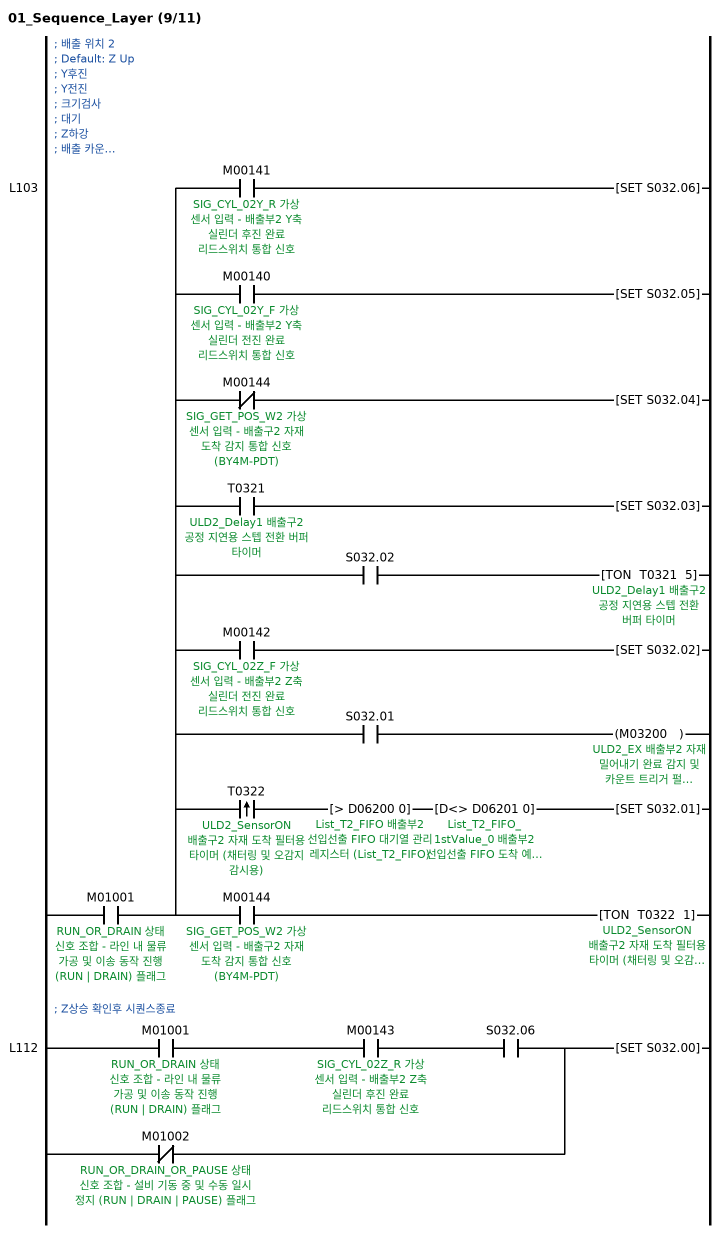
// 
// 배출 위치 2
// 
// Default: Z Up
; L103
LOAD      M01001	// RUN_OR_DRAIN 상태 신호 조합 - 라인 내 물류 가공 및 이송 동작 진행 (RUN | DRAIN) 플래그
MPUSH
AND       M00141	// SIG_CYL_02Y_R 가상 센서 입력 - 배출부2 Y축 실린더 후진 완료 리드스위치 통합 신호
SET       S032.06
MLOAD
AND       M00140	// SIG_CYL_02Y_F 가상 센서 입력 - 배출부2 Y축 실린더 전진 완료 리드스위치 통합 신호
SET       S032.05
MLOAD
AND NOT   M00144	// SIG_GET_POS_W2 가상 센서 입력 - 배출구2 자재 도착 감지 통합 신호 (BY4M-PDT)
SET       S032.04
MLOAD
AND       T0321	// ULD2_Delay1 배출구2 공정 지연용 스텝 전환 버퍼 타이머
SET       S032.03
MLOAD
AND       S032.02
TON       T0321 5	// ULD2_Delay1 배출구2 공정 지연용 스텝 전환 버퍼 타이머
MLOAD
AND       M00142	// SIG_CYL_02Z_F 가상 센서 입력 - 배출부2 Z축 실린더 전진 완료 리드스위치 통합 신호
SET       S032.02
MLOAD
AND       S032.01
OUT       M03200	// ULD2_EX 배출부2 자재 밀어내기 완료 감지 및 카운트 트리거 펄스 (ULD2_EX)
MLOAD
ANDP      T0322	// ULD2_SensorON 배출구2 자재 도착 필터용 타이머 (채터링 및 오감지 감시용)
AND>      D06200 0	// List_T2_FIFO 배출부2 선입선출 FIFO 대기열 관리 레지스터 (List_T2_FIFO)
ANDD<>    D06201 0	// List_T2_FIFO_1stValue_0 배출부2 선입선출 FIFO 도착 예정 시간 데이터 레지스터 하위 16비트 (32비트 연산)
SET       S032.01
MPOP
AND       M00144	// SIG_GET_POS_W2 가상 센서 입력 - 배출구2 자재 도착 감지 통합 신호 (BY4M-PDT)
TON       T0322 1	// ULD2_SensorON 배출구2 자재 도착 필터용 타이머 (채터링 및 오감지 감시용)
// output comment: Y후진
// output comment: Y전진
// output comment: 크기검사
// output comment: 대기
// output comment: Z하강
// output comment: 배출 카운트
// output comment: 도착감지
// output comment: 채터링->데이터오염 방지
; L112
LOAD      M01001	// RUN_OR_DRAIN 상태 신호 조합 - 라인 내 물류 가공 및 이송 동작 진행 (RUN | DRAIN) 플래그
AND       M00143	// SIG_CYL_02Z_R 가상 센서 입력 - 배출부2 Z축 실린더 후진 완료 리드스위치 통합 신호
AND       S032.06
OR NOT    M01002	// RUN_OR_DRAIN_OR_PAUSE 상태 신호 조합 - 설비 기동 중 및 수동 일시 정지 (RUN | DRAIN | PAUSE) 플래그
SET       S032.00
// output comment: Z상승 확인후 시퀀스종료

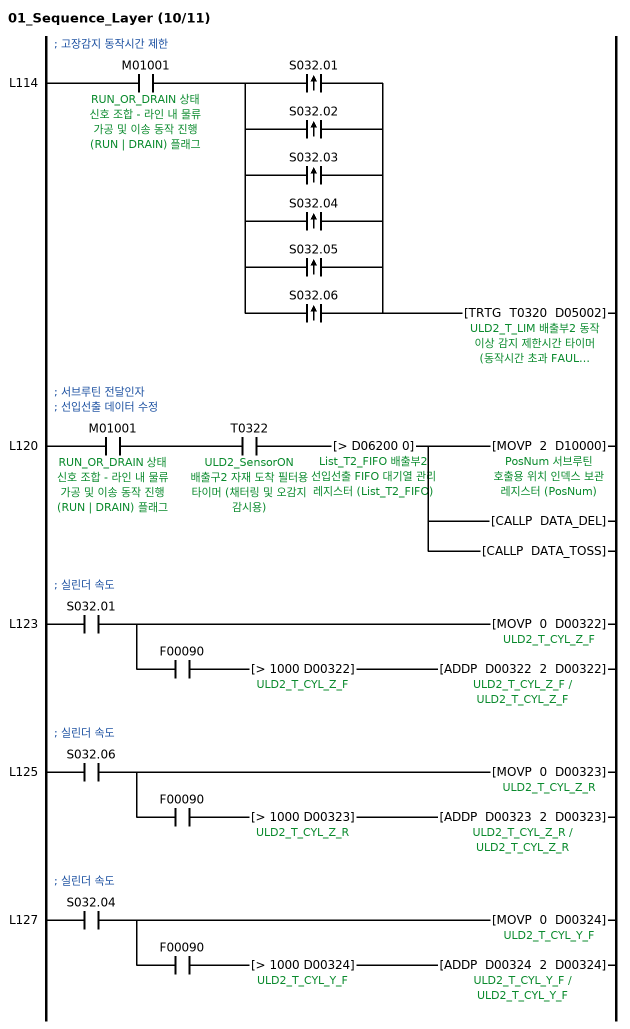
; L114
LOAD      M01001	// RUN_OR_DRAIN 상태 신호 조합 - 라인 내 물류 가공 및 이송 동작 진행 (RUN | DRAIN) 플래그
LOADP     S032.01
ORP       S032.02
ORP       S032.03
ORP       S032.04
ORP       S032.05
ORP       S032.06
AND LOAD
TRTG      T0320 D05002	// ULD2_T_LIM 배출부2 동작 이상 감지 제한시간 타이머 (동작시간 초과 FAULT 트리거) / T_Limit 단위 동작 고장 감지 제한시간(타임아웃) 기준값 설정 레지스터
// output comment: 고장감지 동작시간 제한
; L120
LOAD      M01001	// RUN_OR_DRAIN 상태 신호 조합 - 라인 내 물류 가공 및 이송 동작 진행 (RUN | DRAIN) 플래그
AND       T0322	// ULD2_SensorON 배출구2 자재 도착 필터용 타이머 (채터링 및 오감지 감시용)
AND>      D06200 0	// List_T2_FIFO 배출부2 선입선출 FIFO 대기열 관리 레지스터 (List_T2_FIFO)
MOVP      2 D10000	// PosNum 서브루틴 호출용 위치 인덱스 보관 레지스터 (PosNum)
CALLP     DATA_DEL
CALLP     DATA_TOSS
// output comment: 서브루틴 전달인자
// output comment: 선입선출 데이터 수정
; L123
LOAD      S032.01
MOVP      0 D00322	// ULD2_T_CYL_Z_F
AND       F00090
AND>      1000 D00322	// ULD2_T_CYL_Z_F
ADDP      D00322 2 D00322	// ULD2_T_CYL_Z_F / ULD2_T_CYL_Z_F
// output comment: 실린더 속도
; L125
LOAD      S032.06
MOVP      0 D00323	// ULD2_T_CYL_Z_R
AND       F00090
AND>      1000 D00323	// ULD2_T_CYL_Z_R
ADDP      D00323 2 D00323	// ULD2_T_CYL_Z_R / ULD2_T_CYL_Z_R
// output comment: 실린더 속도
; L127
LOAD      S032.04
MOVP      0 D00324	// ULD2_T_CYL_Y_F
AND       F00090
AND>      1000 D00324	// ULD2_T_CYL_Y_F
ADDP      D00324 2 D00324	// ULD2_T_CYL_Y_F / ULD2_T_CYL_Y_F
// output comment: 실린더 속도

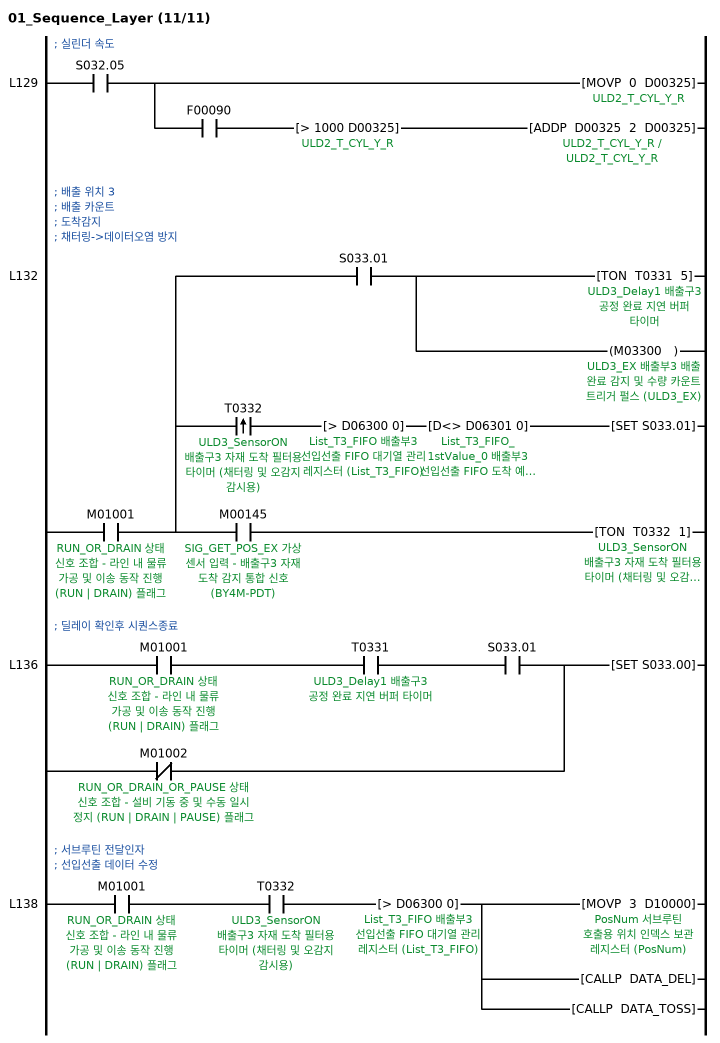
; L129
LOAD      S032.05
MOVP      0 D00325	// ULD2_T_CYL_Y_R
AND       F00090
AND>      1000 D00325	// ULD2_T_CYL_Y_R
ADDP      D00325 2 D00325	// ULD2_T_CYL_Y_R / ULD2_T_CYL_Y_R
// output comment: 실린더 속도
// 배출 위치 3
; L132
LOAD      M01001	// RUN_OR_DRAIN 상태 신호 조합 - 라인 내 물류 가공 및 이송 동작 진행 (RUN | DRAIN) 플래그
MPUSH
AND       S033.01
TON       T0331 5	// ULD3_Delay1 배출구3 공정 완료 지연 버퍼 타이머
OUT       M03300	// ULD3_EX 배출부3 배출 완료 감지 및 수량 카운트 트리거 펄스 (ULD3_EX)
MLOAD
ANDP      T0332	// ULD3_SensorON 배출구3 자재 도착 필터용 타이머 (채터링 및 오감지 감시용)
AND>      D06300 0	// List_T3_FIFO 배출부3 선입선출 FIFO 대기열 관리 레지스터 (List_T3_FIFO)
ANDD<>    D06301 0	// List_T3_FIFO_1stValue_0 배출부3 선입선출 FIFO 도착 예정 시간 데이터 레지스터 하위 16비트 (32비트 연산)
SET       S033.01
MPOP
AND       M00145	// SIG_GET_POS_EX 가상 센서 입력 - 배출구3 자재 도착 감지 통합 신호 (BY4M-PDT)
TON       T0332 1	// ULD3_SensorON 배출구3 자재 도착 필터용 타이머 (채터링 및 오감지 감시용)
// output comment: 배출 카운트
// output comment: 도착감지
// output comment: 채터링->데이터오염 방지
; L136
LOAD      M01001	// RUN_OR_DRAIN 상태 신호 조합 - 라인 내 물류 가공 및 이송 동작 진행 (RUN | DRAIN) 플래그
AND       T0331	// ULD3_Delay1 배출구3 공정 완료 지연 버퍼 타이머
AND       S033.01
OR NOT    M01002	// RUN_OR_DRAIN_OR_PAUSE 상태 신호 조합 - 설비 기동 중 및 수동 일시 정지 (RUN | DRAIN | PAUSE) 플래그
SET       S033.00
// output comment: 딜레이 확인후 시퀀스종료
; L138
LOAD      M01001	// RUN_OR_DRAIN 상태 신호 조합 - 라인 내 물류 가공 및 이송 동작 진행 (RUN | DRAIN) 플래그
AND       T0332	// ULD3_SensorON 배출구3 자재 도착 필터용 타이머 (채터링 및 오감지 감시용)
AND>      D06300 0	// List_T3_FIFO 배출부3 선입선출 FIFO 대기열 관리 레지스터 (List_T3_FIFO)
MOVP      3 D10000	// PosNum 서브루틴 호출용 위치 인덱스 보관 레지스터 (PosNum)
CALLP     DATA_DEL
CALLP     DATA_TOSS
// output comment: 서브루틴 전달인자
// output comment: 선입선출 데이터 수정

PROGRAM 97_Error_Layer (task: 스캔 프로그램)

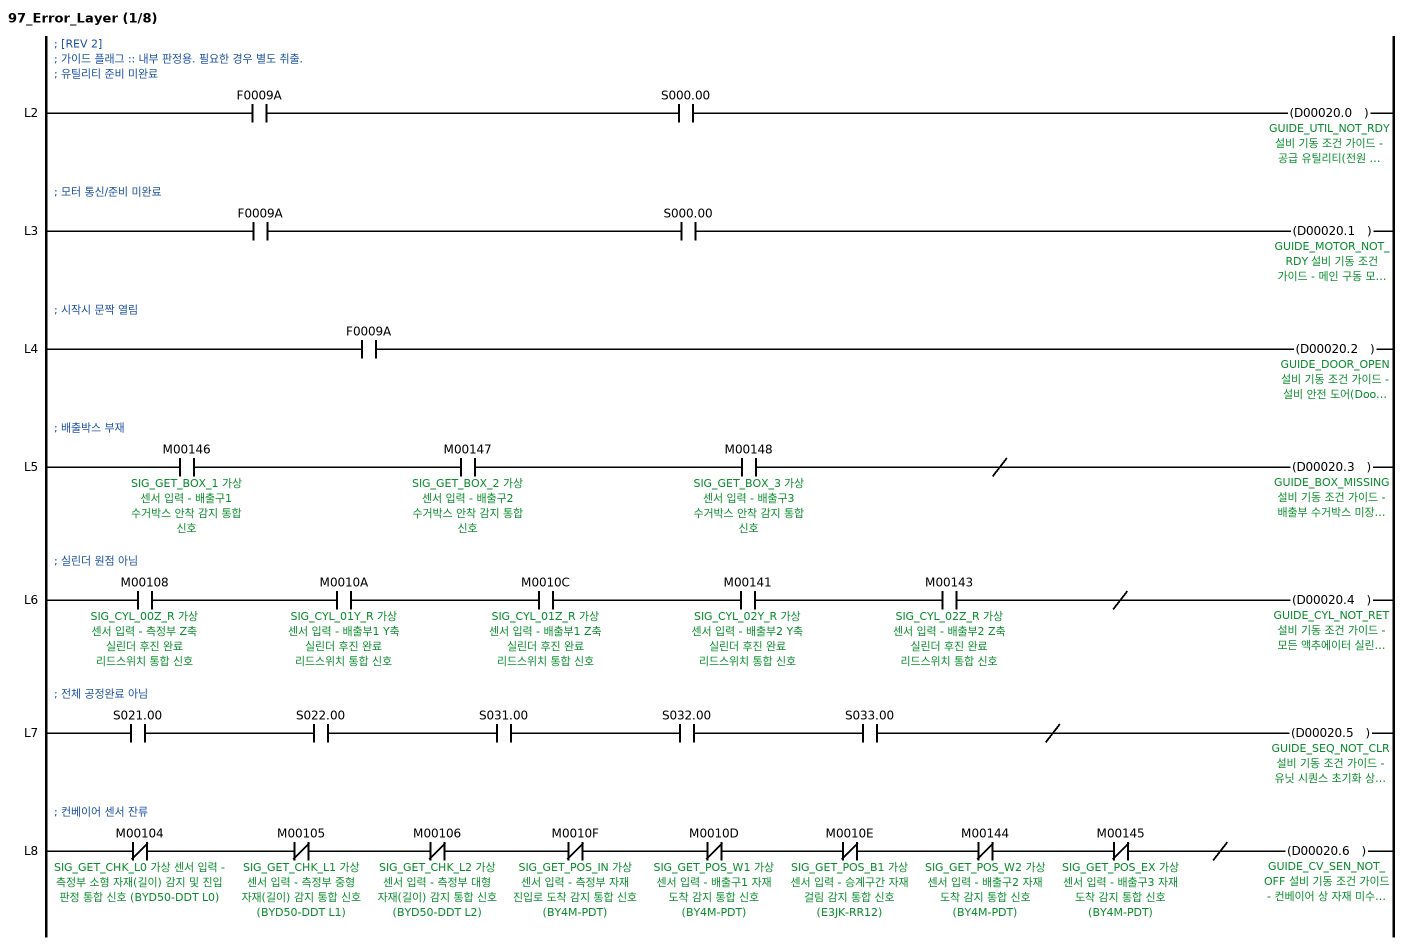
// [REV 2]
// 가이드 플래그 :: 내부 판정용. 필요한 경우 별도 취출.
; L2
LOAD      F0009A
AND       S000.00
OUT       D00020.0	// GUIDE_UTIL_NOT_RDY 설비 기동 조건 가이드 - 공급 유틸리티(전원 및 공압) 공급 상태 미완료 감지 가이드 비트
// output comment: 유틸리티 준비 미완료
; L3
LOAD      F0009A
AND       S000.00
OUT       D00020.1	// GUIDE_MOTOR_NOT_RDY 설비 기동 조건 가이드 - 메인 구동 모터 드라이버 통신 및 준비 상태 미완료 감지 가이드 비트
// output comment: 모터 통신/준비 미완료
; L4
LOAD      F0009A
OUT       D00020.2	// GUIDE_DOOR_OPEN 설비 기동 조건 가이드 - 설비 안전 도어(Door Interface) 개방 상태 감지 가이드 비트
// output comment: 시작시 문짝 열림
; L5
LOAD      M00146	// SIG_GET_BOX_1 가상 센서 입력 - 배출구1 수거박스 안착 감지 통합 신호
AND       M00147	// SIG_GET_BOX_2 가상 센서 입력 - 배출구2 수거박스 안착 감지 통합 신호
AND       M00148	// SIG_GET_BOX_3 가상 센서 입력 - 배출구3 수거박스 안착 감지 통합 신호
NOT
OUT       D00020.3	// GUIDE_BOX_MISSING 설비 기동 조건 가이드 - 배출부 수거박스 미장착 감지 가이드 비트
// output comment: 배출박스 부재
; L6
LOAD      M00108	// SIG_CYL_00Z_R 가상 센서 입력 - 측정부 Z축 실린더 후진 완료 리드스위치 통합 신호
AND       M0010A	// SIG_CYL_01Y_R 가상 센서 입력 - 배출부1 Y축 실린더 후진 완료 리드스위치 통합 신호
AND       M0010C	// SIG_CYL_01Z_R 가상 센서 입력 - 배출부1 Z축 실린더 후진 완료 리드스위치 통합 신호
AND       M00141	// SIG_CYL_02Y_R 가상 센서 입력 - 배출부2 Y축 실린더 후진 완료 리드스위치 통합 신호
AND       M00143	// SIG_CYL_02Z_R 가상 센서 입력 - 배출부2 Z축 실린더 후진 완료 리드스위치 통합 신호
NOT
OUT       D00020.4	// GUIDE_CYL_NOT_RET 설비 기동 조건 가이드 - 모든 액추에이터 실린더 원점(후퇴) 미복귀 가이드 비트
// output comment: 실린더 원점 아님
; L7
LOAD      S021.00
AND       S022.00
AND       S031.00
AND       S032.00
AND       S033.00
NOT
OUT       D00020.5	// GUIDE_SEQ_NOT_CLR 설비 기동 조건 가이드 - 유닛 시퀀스 초기화 상태 미복귀 가이드 비트
// output comment: 전체 공정완료 아님
; L8
LOAD NOT  M00104	// SIG_GET_CHK_L0 가상 센서 입력 - 측정부 소형 자재(길이) 감지 및 진입 판정 통합 신호 (BYD50-DDT L0)
AND NOT   M00105	// SIG_GET_CHK_L1 가상 센서 입력 - 측정부 중형 자재(길이) 감지 통합 신호 (BYD50-DDT L1)
AND NOT   M00106	// SIG_GET_CHK_L2 가상 센서 입력 - 측정부 대형 자재(길이) 감지 통합 신호 (BYD50-DDT L2)
AND NOT   M0010F	// SIG_GET_POS_IN 가상 센서 입력 - 측정부 자재 진입로 도착 감지 통합 신호 (BY4M-PDT)
AND NOT   M0010D	// SIG_GET_POS_W1 가상 센서 입력 - 배출구1 자재 도착 감지 통합 신호 (BY4M-PDT)
AND NOT   M0010E	// SIG_GET_POS_B1 가상 센서 입력 - 승계구간 자재 걸림 감지 통합 신호 (E3JK-RR12)
AND NOT   M00144	// SIG_GET_POS_W2 가상 센서 입력 - 배출구2 자재 도착 감지 통합 신호 (BY4M-PDT)
AND NOT   M00145	// SIG_GET_POS_EX 가상 센서 입력 - 배출구3 자재 도착 감지 통합 신호 (BY4M-PDT)
NOT
OUT       D00020.6	// GUIDE_CV_SEN_NOT_OFF 설비 기동 조건 가이드 - 컨베이어 상 자재 미수거 잔류 감지 가이드 비트
// output comment: 컨베이어 센서 잔류

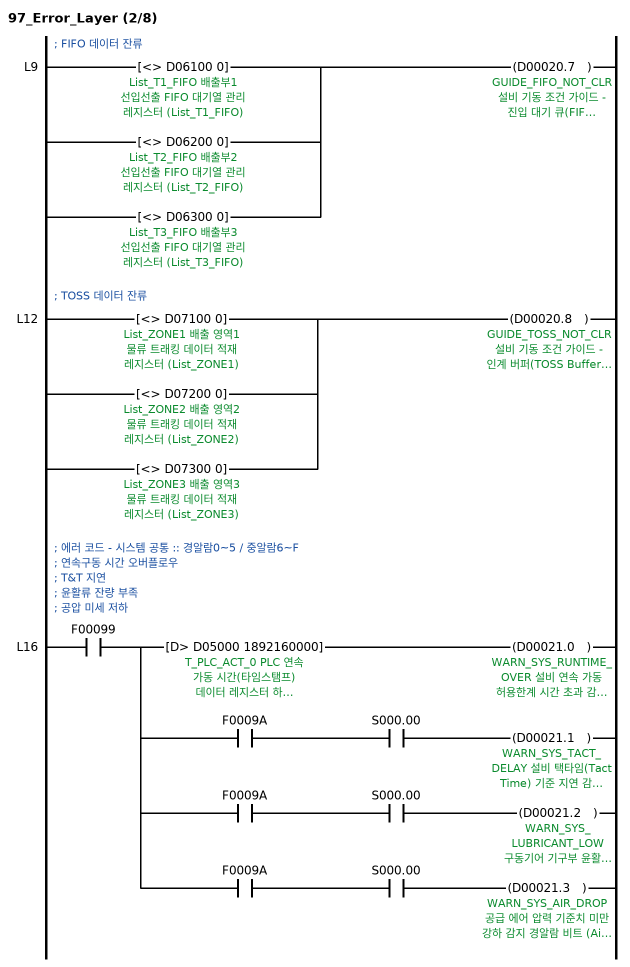
; L9
LOAD<>    D06100 0	// List_T1_FIFO 배출부1 선입선출 FIFO 대기열 관리 레지스터 (List_T1_FIFO)
OR<>      D06200 0	// List_T2_FIFO 배출부2 선입선출 FIFO 대기열 관리 레지스터 (List_T2_FIFO)
OR<>      D06300 0	// List_T3_FIFO 배출부3 선입선출 FIFO 대기열 관리 레지스터 (List_T3_FIFO)
OUT       D00020.7	// GUIDE_FIFO_NOT_CLR 설비 기동 조건 가이드 - 진입 대기 큐(FIFO Queue) 잔류 데이터 존재 가이드 비트
// output comment: FIFO 데이터 잔류
; L12
LOAD<>    D07100 0	// List_ZONE1 배출 영역1 물류 트래킹 데이터 적재 레지스터 (List_ZONE1)
OR<>      D07200 0	// List_ZONE2 배출 영역2 물류 트래킹 데이터 적재 레지스터 (List_ZONE2)
OR<>      D07300 0	// List_ZONE3 배출 영역3 물류 트래킹 데이터 적재 레지스터 (List_ZONE3)
OUT       D00020.8	// GUIDE_TOSS_NOT_CLR 설비 기동 조건 가이드 - 인계 버퍼(TOSS Buffer) 잔류 데이터 존재 가이드 비트
// output comment: TOSS 데이터 잔류
// 에러 코드 - 시스템 공통 :: 경알람0~5 / 중알람6~F
; L16
LOAD      F00099
MPUSH
ANDD>     D05000 1892160000	// T_PLC_ACT_0 PLC 연속 가동 시간(타임스탬프) 데이터 레지스터 하위 16비트 (0.1초 해상도)
OUT       D00021.0	// WARN_SYS_RUNTIME_OVER 설비 연속 가동 허용한계 시간 초과 감지 경알람 비트 (교대 가동 관리)
MLOAD
AND       F0009A
AND       S000.00
OUT       D00021.1	// WARN_SYS_TACT_DELAY 설비 택타임(Tact Time) 기준 지연 감지 경알람 비트 (기구 마모/노후 감시)
MLOAD
AND       F0009A
AND       S000.00
OUT       D00021.2	// WARN_SYS_LUBRICANT_LOW 구동기어 기구부 윤활유 레벨 기준치 미만 저하 감지 경알람 비트 (Oil Low)
MPOP
AND       F0009A
AND       S000.00
OUT       D00021.3	// WARN_SYS_AIR_DROP 공급 에어 압력 기준치 미만 강하 감지 경알람 비트 (Air Leak)
// output comment: 연속구동 시간 오버플로우
// output comment: T&T 지연
// output comment: 윤활류 잔량 부족
// output comment: 공압 미세 저하

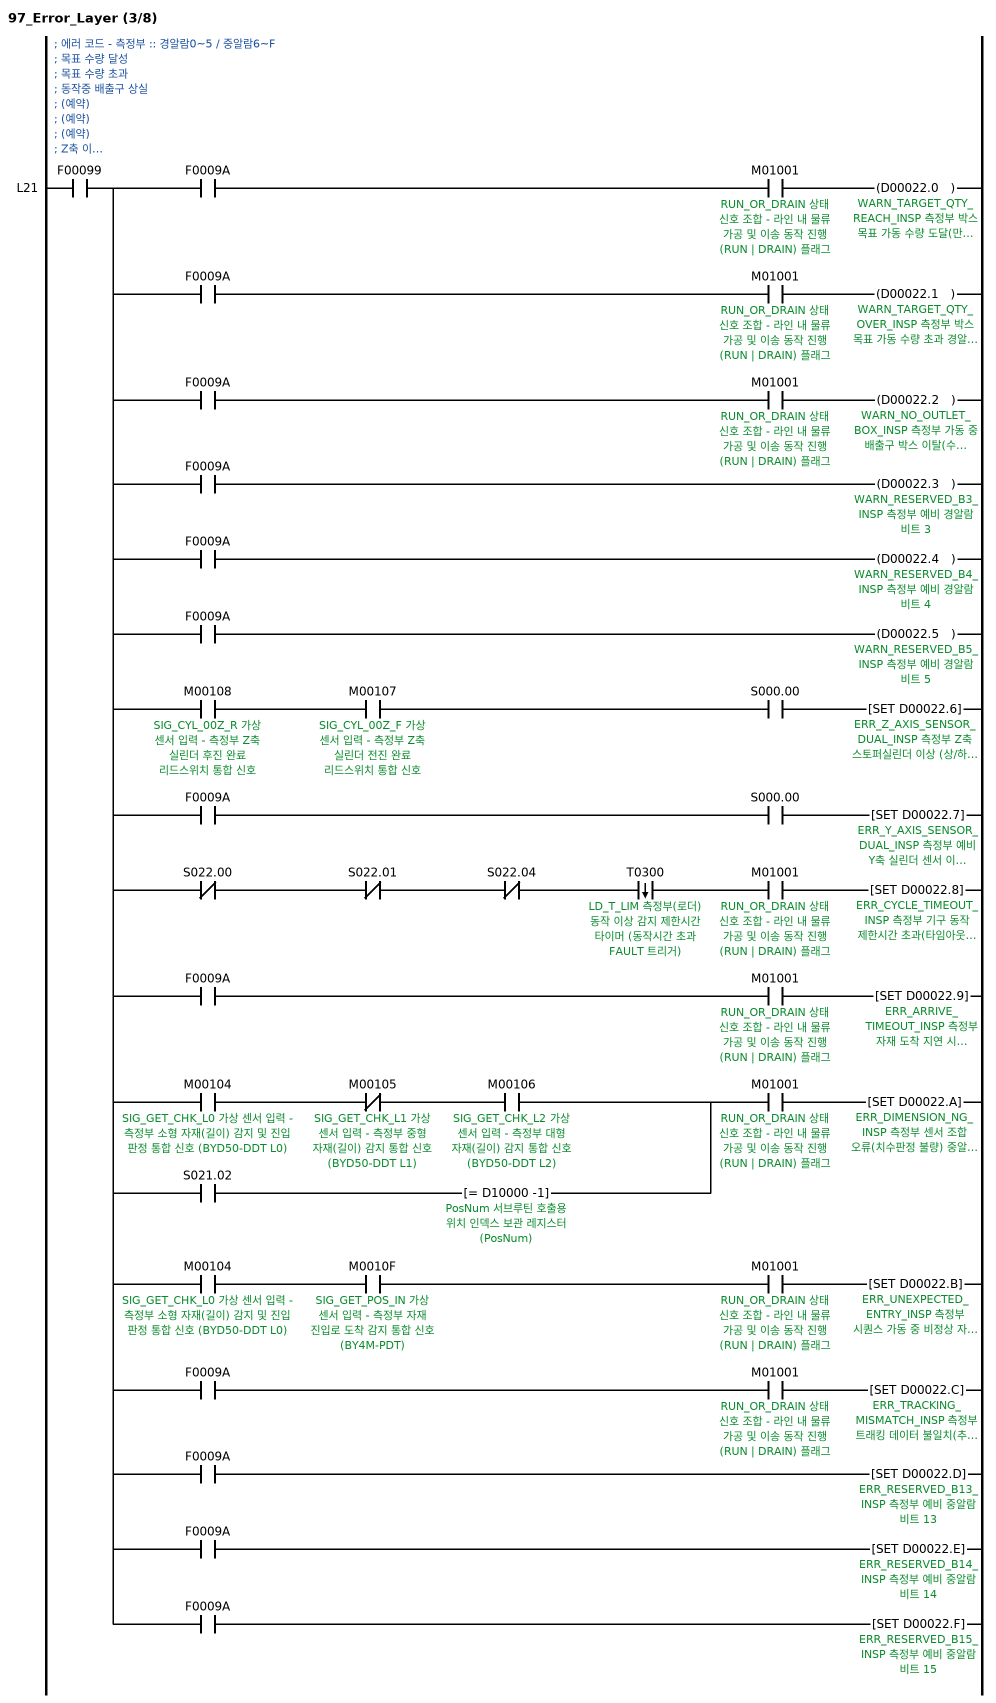
// 에러 코드 - 측정부 :: 경알람0~5 / 중알람6~F
; L21
LOAD      F00099
MPUSH
AND       F0009A
AND       M01001	// RUN_OR_DRAIN 상태 신호 조합 - 라인 내 물류 가공 및 이송 동작 진행 (RUN | DRAIN) 플래그
OUT       D00022.0	// WARN_TARGET_QTY_REACH_INSP 측정부 박스 목표 가동 수량 도달(만재 상태) 경알람 비트
MLOAD
AND       F0009A
AND       M01001	// RUN_OR_DRAIN 상태 신호 조합 - 라인 내 물류 가공 및 이송 동작 진행 (RUN | DRAIN) 플래그
OUT       D00022.1	// WARN_TARGET_QTY_OVER_INSP 측정부 박스 목표 가동 수량 초과 경알람 비트
MLOAD
AND       F0009A
AND       M01001	// RUN_OR_DRAIN 상태 신호 조합 - 라인 내 물류 가공 및 이송 동작 진행 (RUN | DRAIN) 플래그
OUT       D00022.2	// WARN_NO_OUTLET_BOX_INSP 측정부 가동 중 배출구 박스 이탈(수거 상실) 경알람 비트
MLOAD
AND       F0009A
OUT       D00022.3	// WARN_RESERVED_B3_INSP 측정부 예비 경알람 비트 3
MLOAD
AND       F0009A
OUT       D00022.4	// WARN_RESERVED_B4_INSP 측정부 예비 경알람 비트 4
MLOAD
AND       F0009A
OUT       D00022.5	// WARN_RESERVED_B5_INSP 측정부 예비 경알람 비트 5
MLOAD
AND       M00108	// SIG_CYL_00Z_R 가상 센서 입력 - 측정부 Z축 실린더 후진 완료 리드스위치 통합 신호
AND       M00107	// SIG_CYL_00Z_F 가상 센서 입력 - 측정부 Z축 실린더 전진 완료 리드스위치 통합 신호
AND       S000.00
SET       D00022.6	// ERR_Z_AXIS_SENSOR_DUAL_INSP 측정부 Z축 스토퍼실린더 이상 (상/하한 센서 동시 ON) 중알람 비트
MLOAD
AND       F0009A
AND       S000.00
SET       D00022.7	// ERR_Y_AXIS_SENSOR_DUAL_INSP 측정부 예비 Y축 실린더 센서 이상 중알람 비트 7
MLOAD
AND NOT   S022.00
AND NOT   S022.01
AND NOT   S022.04
ANDN      T0300	// LD_T_LIM 측정부(로더) 동작 이상 감지 제한시간 타이머 (동작시간 초과 FAULT 트리거)
AND       M01001	// RUN_OR_DRAIN 상태 신호 조합 - 라인 내 물류 가공 및 이송 동작 진행 (RUN | DRAIN) 플래그
SET       D00022.8	// ERR_CYCLE_TIMEOUT_INSP 측정부 기구 동작 제한시간 초과(타임아웃) 중알람 비트
MLOAD
AND       F0009A
AND       M01001	// RUN_OR_DRAIN 상태 신호 조합 - 라인 내 물류 가공 및 이송 동작 진행 (RUN | DRAIN) 플래그
SET       D00022.9	// ERR_ARRIVE_TIMEOUT_INSP 측정부 자재 도착 지연 시간 초과(FIFO 대기시간 초과) 중알람 비트
MLOAD
LOAD      M00104	// SIG_GET_CHK_L0 가상 센서 입력 - 측정부 소형 자재(길이) 감지 및 진입 판정 통합 신호 (BYD50-DDT L0)
AND NOT   M00105	// SIG_GET_CHK_L1 가상 센서 입력 - 측정부 중형 자재(길이) 감지 통합 신호 (BYD50-DDT L1)
AND       M00106	// SIG_GET_CHK_L2 가상 센서 입력 - 측정부 대형 자재(길이) 감지 통합 신호 (BYD50-DDT L2)
LOAD      S021.02
AND=      D10000 -1	// PosNum 서브루틴 호출용 위치 인덱스 보관 레지스터 (PosNum)
OR LOAD
AND LOAD
AND       M01001	// RUN_OR_DRAIN 상태 신호 조합 - 라인 내 물류 가공 및 이송 동작 진행 (RUN | DRAIN) 플래그
SET       D00022.A	// ERR_DIMENSION_NG_INSP 측정부 센서 조합 오류(치수판정 불량) 중알람 비트
MLOAD
AND       M00104	// SIG_GET_CHK_L0 가상 센서 입력 - 측정부 소형 자재(길이) 감지 및 진입 판정 통합 신호 (BYD50-DDT L0)
AND       M0010F	// SIG_GET_POS_IN 가상 센서 입력 - 측정부 자재 진입로 도착 감지 통합 신호 (BY4M-PDT)
AND       M01001	// RUN_OR_DRAIN 상태 신호 조합 - 라인 내 물류 가공 및 이송 동작 진행 (RUN | DRAIN) 플래그
SET       D00022.B	// ERR_UNEXPECTED_ENTRY_INSP 측정부 시퀀스 가동 중 비정상 자재 진입 중알람 비트
MLOAD
AND       F0009A
AND       M01001	// RUN_OR_DRAIN 상태 신호 조합 - 라인 내 물류 가공 및 이송 동작 진행 (RUN | DRAIN) 플래그
SET       D00022.C	// ERR_TRACKING_MISMATCH_INSP 측정부 트래킹 데이터 불일치(추적 오동작) 중알람 비트
MLOAD
AND       F0009A
SET       D00022.D	// ERR_RESERVED_B13_INSP 측정부 예비 중알람 비트 13
MLOAD
AND       F0009A
SET       D00022.E	// ERR_RESERVED_B14_INSP 측정부 예비 중알람 비트 14
MPOP
AND       F0009A
SET       D00022.F	// ERR_RESERVED_B15_INSP 측정부 예비 중알람 비트 15
// output comment: 목표 수량 달성
// output comment: 목표 수량 초과
// output comment: 동작중 배출구 상실
// output comment: (예약)
// output comment: (예약)
// output comment: (예약)
// output comment: Z축 이상
// output comment: Y축 이상
// output comment: 동작시간 초과
// output comment: 도착시간 초과
// output comment: 치수판정 불량
// output comment: 작동중 투입
// output comment: 추적 불일치
// output comment: (예약)
// output comment: (예약)
// output comment: (예약)

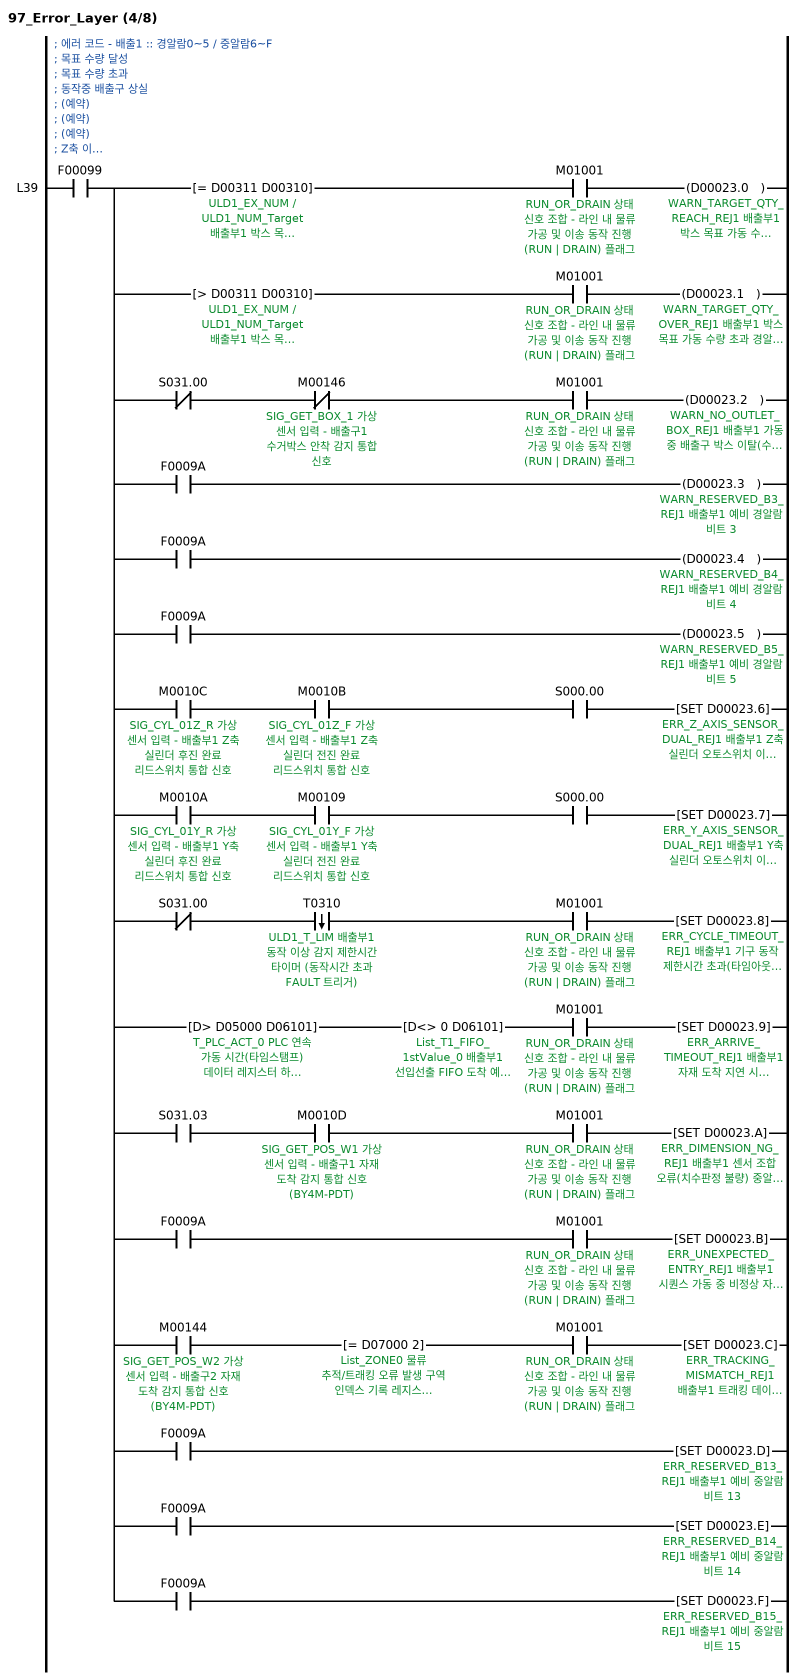
// 에러 코드 - 배출1 :: 경알람0~5 / 중알람6~F
; L39
LOAD      F00099
MPUSH
AND=      D00311 D00310	// ULD1_EX_NUM / ULD1_NUM_Target 배출부1 박스 목표 분류/배출 완료 수량 레지스터
AND       M01001	// RUN_OR_DRAIN 상태 신호 조합 - 라인 내 물류 가공 및 이송 동작 진행 (RUN | DRAIN) 플래그
OUT       D00023.0	// WARN_TARGET_QTY_REACH_REJ1 배출부1 박스 목표 가동 수량 도달(만재 상태) 경알람 비트
MLOAD
AND>      D00311 D00310	// ULD1_EX_NUM / ULD1_NUM_Target 배출부1 박스 목표 분류/배출 완료 수량 레지스터
AND       M01001	// RUN_OR_DRAIN 상태 신호 조합 - 라인 내 물류 가공 및 이송 동작 진행 (RUN | DRAIN) 플래그
OUT       D00023.1	// WARN_TARGET_QTY_OVER_REJ1 배출부1 박스 목표 가동 수량 초과 경알람 비트
MLOAD
AND NOT   S031.00
AND NOT   M00146	// SIG_GET_BOX_1 가상 센서 입력 - 배출구1 수거박스 안착 감지 통합 신호
AND       M01001	// RUN_OR_DRAIN 상태 신호 조합 - 라인 내 물류 가공 및 이송 동작 진행 (RUN | DRAIN) 플래그
OUT       D00023.2	// WARN_NO_OUTLET_BOX_REJ1 배출부1 가동 중 배출구 박스 이탈(수거 상실) 경알람 비트
MLOAD
AND       F0009A
OUT       D00023.3	// WARN_RESERVED_B3_REJ1 배출부1 예비 경알람 비트 3
MLOAD
AND       F0009A
OUT       D00023.4	// WARN_RESERVED_B4_REJ1 배출부1 예비 경알람 비트 4
MLOAD
AND       F0009A
OUT       D00023.5	// WARN_RESERVED_B5_REJ1 배출부1 예비 경알람 비트 5
MLOAD
AND       M0010C	// SIG_CYL_01Z_R 가상 센서 입력 - 배출부1 Z축 실린더 후진 완료 리드스위치 통합 신호
AND       M0010B	// SIG_CYL_01Z_F 가상 센서 입력 - 배출부1 Z축 실린더 전진 완료 리드스위치 통합 신호
AND       S000.00
SET       D00023.6	// ERR_Z_AXIS_SENSOR_DUAL_REJ1 배출부1 Z축 실린더 오토스위치 이상 (상/하한 센서 동시 ON) 중알람 비트
MLOAD
AND       M0010A	// SIG_CYL_01Y_R 가상 센서 입력 - 배출부1 Y축 실린더 후진 완료 리드스위치 통합 신호
AND       M00109	// SIG_CYL_01Y_F 가상 센서 입력 - 배출부1 Y축 실린더 전진 완료 리드스위치 통합 신호
AND       S000.00
SET       D00023.7	// ERR_Y_AXIS_SENSOR_DUAL_REJ1 배출부1 Y축 실린더 오토스위치 이상 (전/후진 센서 동시 ON) 중알람 비트
MLOAD
AND NOT   S031.00
ANDN      T0310	// ULD1_T_LIM 배출부1 동작 이상 감지 제한시간 타이머 (동작시간 초과 FAULT 트리거)
AND       M01001	// RUN_OR_DRAIN 상태 신호 조합 - 라인 내 물류 가공 및 이송 동작 진행 (RUN | DRAIN) 플래그
SET       D00023.8	// ERR_CYCLE_TIMEOUT_REJ1 배출부1 기구 동작 제한시간 초과(타임아웃) 중알람 비트
MLOAD
ANDD>     D05000 D06101	// T_PLC_ACT_0 PLC 연속 가동 시간(타임스탬프) 데이터 레지스터 하위 16비트 (0.1초 해상도) / List_T1_FIFO_1stValue_0 배출부1 선입선출 FIFO 도착 예정 시간 데이터 레지스터 하위 16비트 (32비트 연산)
ANDD<>    0 D06101	// List_T1_FIFO_1stValue_0 배출부1 선입선출 FIFO 도착 예정 시간 데이터 레지스터 하위 16비트 (32비트 연산)
AND       M01001	// RUN_OR_DRAIN 상태 신호 조합 - 라인 내 물류 가공 및 이송 동작 진행 (RUN | DRAIN) 플래그
SET       D00023.9	// ERR_ARRIVE_TIMEOUT_REJ1 배출부1 자재 도착 지연 시간 초과(FIFO 대기시간 초과) 중알람 비트
MLOAD
AND       S031.03
AND       M0010D	// SIG_GET_POS_W1 가상 센서 입력 - 배출구1 자재 도착 감지 통합 신호 (BY4M-PDT)
AND       M01001	// RUN_OR_DRAIN 상태 신호 조합 - 라인 내 물류 가공 및 이송 동작 진행 (RUN | DRAIN) 플래그
SET       D00023.A	// ERR_DIMENSION_NG_REJ1 배출부1 센서 조합 오류(치수판정 불량) 중알람 비트
MLOAD
AND       F0009A
AND       M01001	// RUN_OR_DRAIN 상태 신호 조합 - 라인 내 물류 가공 및 이송 동작 진행 (RUN | DRAIN) 플래그
SET       D00023.B	// ERR_UNEXPECTED_ENTRY_REJ1 배출부1 시퀀스 가동 중 비정상 자재 진입 중알람 비트
MLOAD
AND       M00144	// SIG_GET_POS_W2 가상 센서 입력 - 배출구2 자재 도착 감지 통합 신호 (BY4M-PDT)
AND=      D07000 2	// List_ZONE0 물류 추적/트래킹 오류 발생 구역 인덱스 기록 레지스터 (List_ZONE0)
AND       M01001	// RUN_OR_DRAIN 상태 신호 조합 - 라인 내 물류 가공 및 이송 동작 진행 (RUN | DRAIN) 플래그
SET       D00023.C	// ERR_TRACKING_MISMATCH_REJ1 배출부1 트래킹 데이터 불일치(추적 오동작) 중알람 비트
MLOAD
AND       F0009A
SET       D00023.D	// ERR_RESERVED_B13_REJ1 배출부1 예비 중알람 비트 13
MLOAD
AND       F0009A
SET       D00023.E	// ERR_RESERVED_B14_REJ1 배출부1 예비 중알람 비트 14
MPOP
AND       F0009A
SET       D00023.F	// ERR_RESERVED_B15_REJ1 배출부1 예비 중알람 비트 15
// output comment: 목표 수량 달성
// output comment: 목표 수량 초과
// output comment: 동작중 배출구 상실
// output comment: (예약)
// output comment: (예약)
// output comment: (예약)
// output comment: Z축 이상
// output comment: Y축 이상
// output comment: 동작시간 초과
// output comment: 도착시간 초과
// output comment: 치수판정 불량
// output comment: 작동중 투입
// output comment: 추적 불일치
// output comment: (예약)
// output comment: (예약)
// output comment: (예약)

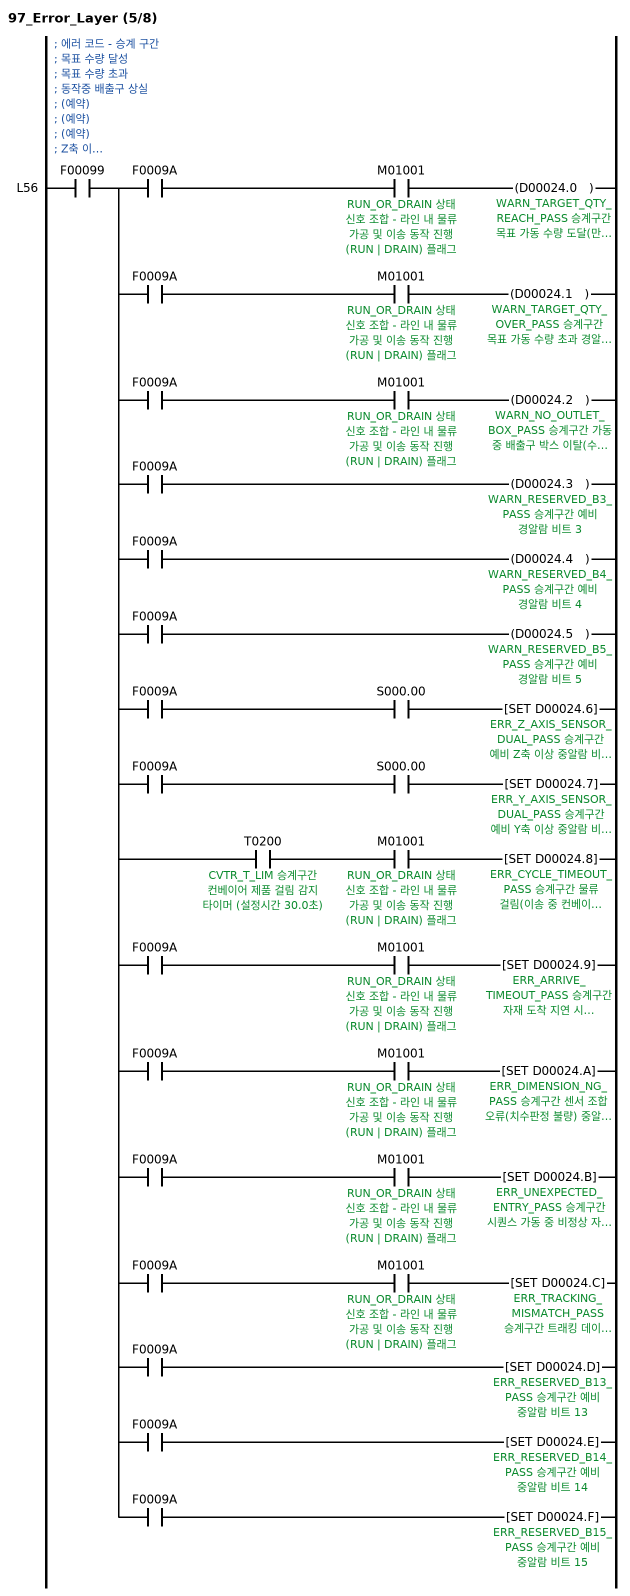
// 에러 코드 - 승계 구간
; L56
LOAD      F00099
MPUSH
AND       F0009A
AND       M01001	// RUN_OR_DRAIN 상태 신호 조합 - 라인 내 물류 가공 및 이송 동작 진행 (RUN | DRAIN) 플래그
OUT       D00024.0	// WARN_TARGET_QTY_REACH_PASS 승계구간 목표 가동 수량 도달(만재 상태) 경알람 비트
MLOAD
AND       F0009A
AND       M01001	// RUN_OR_DRAIN 상태 신호 조합 - 라인 내 물류 가공 및 이송 동작 진행 (RUN | DRAIN) 플래그
OUT       D00024.1	// WARN_TARGET_QTY_OVER_PASS 승계구간 목표 가동 수량 초과 경알람 비트
MLOAD
AND       F0009A
AND       M01001	// RUN_OR_DRAIN 상태 신호 조합 - 라인 내 물류 가공 및 이송 동작 진행 (RUN | DRAIN) 플래그
OUT       D00024.2	// WARN_NO_OUTLET_BOX_PASS 승계구간 가동 중 배출구 박스 이탈(수거 상실) 경알람 비트
MLOAD
AND       F0009A
OUT       D00024.3	// WARN_RESERVED_B3_PASS 승계구간 예비 경알람 비트 3
MLOAD
AND       F0009A
OUT       D00024.4	// WARN_RESERVED_B4_PASS 승계구간 예비 경알람 비트 4
MLOAD
AND       F0009A
OUT       D00024.5	// WARN_RESERVED_B5_PASS 승계구간 예비 경알람 비트 5
MLOAD
AND       F0009A
AND       S000.00
SET       D00024.6	// ERR_Z_AXIS_SENSOR_DUAL_PASS 승계구간 예비 Z축 이상 중알람 비트 6
MLOAD
AND       F0009A
AND       S000.00
SET       D00024.7	// ERR_Y_AXIS_SENSOR_DUAL_PASS 승계구간 예비 Y축 이상 중알람 비트 7
MLOAD
AND       T0200	// CVTR_T_LIM 승계구간 컨베이어 제품 걸림 감지 타이머 (설정시간 30.0초)
AND       M01001	// RUN_OR_DRAIN 상태 신호 조합 - 라인 내 물류 가공 및 이송 동작 진행 (RUN | DRAIN) 플래그
SET       D00024.8	// ERR_CYCLE_TIMEOUT_PASS 승계구간 물류 걸림(이송 중 컨베이어 지연) 중알람 비트
MLOAD
AND       F0009A
AND       M01001	// RUN_OR_DRAIN 상태 신호 조합 - 라인 내 물류 가공 및 이송 동작 진행 (RUN | DRAIN) 플래그
SET       D00024.9	// ERR_ARRIVE_TIMEOUT_PASS 승계구간 자재 도착 지연 시간 초과(FIFO 대기시간 초과) 중알람 비트
MLOAD
AND       F0009A
AND       M01001	// RUN_OR_DRAIN 상태 신호 조합 - 라인 내 물류 가공 및 이송 동작 진행 (RUN | DRAIN) 플래그
SET       D00024.A	// ERR_DIMENSION_NG_PASS 승계구간 센서 조합 오류(치수판정 불량) 중알람 비트
MLOAD
AND       F0009A
AND       M01001	// RUN_OR_DRAIN 상태 신호 조합 - 라인 내 물류 가공 및 이송 동작 진행 (RUN | DRAIN) 플래그
SET       D00024.B	// ERR_UNEXPECTED_ENTRY_PASS 승계구간 시퀀스 가동 중 비정상 자재 진입 중알람 비트
MLOAD
AND       F0009A
AND       M01001	// RUN_OR_DRAIN 상태 신호 조합 - 라인 내 물류 가공 및 이송 동작 진행 (RUN | DRAIN) 플래그
SET       D00024.C	// ERR_TRACKING_MISMATCH_PASS 승계구간 트래킹 데이터 불일치(추적 오동작) 중알람 비트
MLOAD
AND       F0009A
SET       D00024.D	// ERR_RESERVED_B13_PASS 승계구간 예비 중알람 비트 13
MLOAD
AND       F0009A
SET       D00024.E	// ERR_RESERVED_B14_PASS 승계구간 예비 중알람 비트 14
MPOP
AND       F0009A
SET       D00024.F	// ERR_RESERVED_B15_PASS 승계구간 예비 중알람 비트 15
// output comment: 목표 수량 달성
// output comment: 목표 수량 초과
// output comment: 동작중 배출구 상실
// output comment: (예약)
// output comment: (예약)
// output comment: (예약)
// output comment: Z축 이상
// output comment: Y축 이상
// output comment: 동작시간 초과
// output comment: 도착시간 초과
// output comment: 치수판정 불량
// output comment: 작동중 투입
// output comment: 추적 불일치
// output comment: (예약)
// output comment: (예약)
// output comment: (예약)

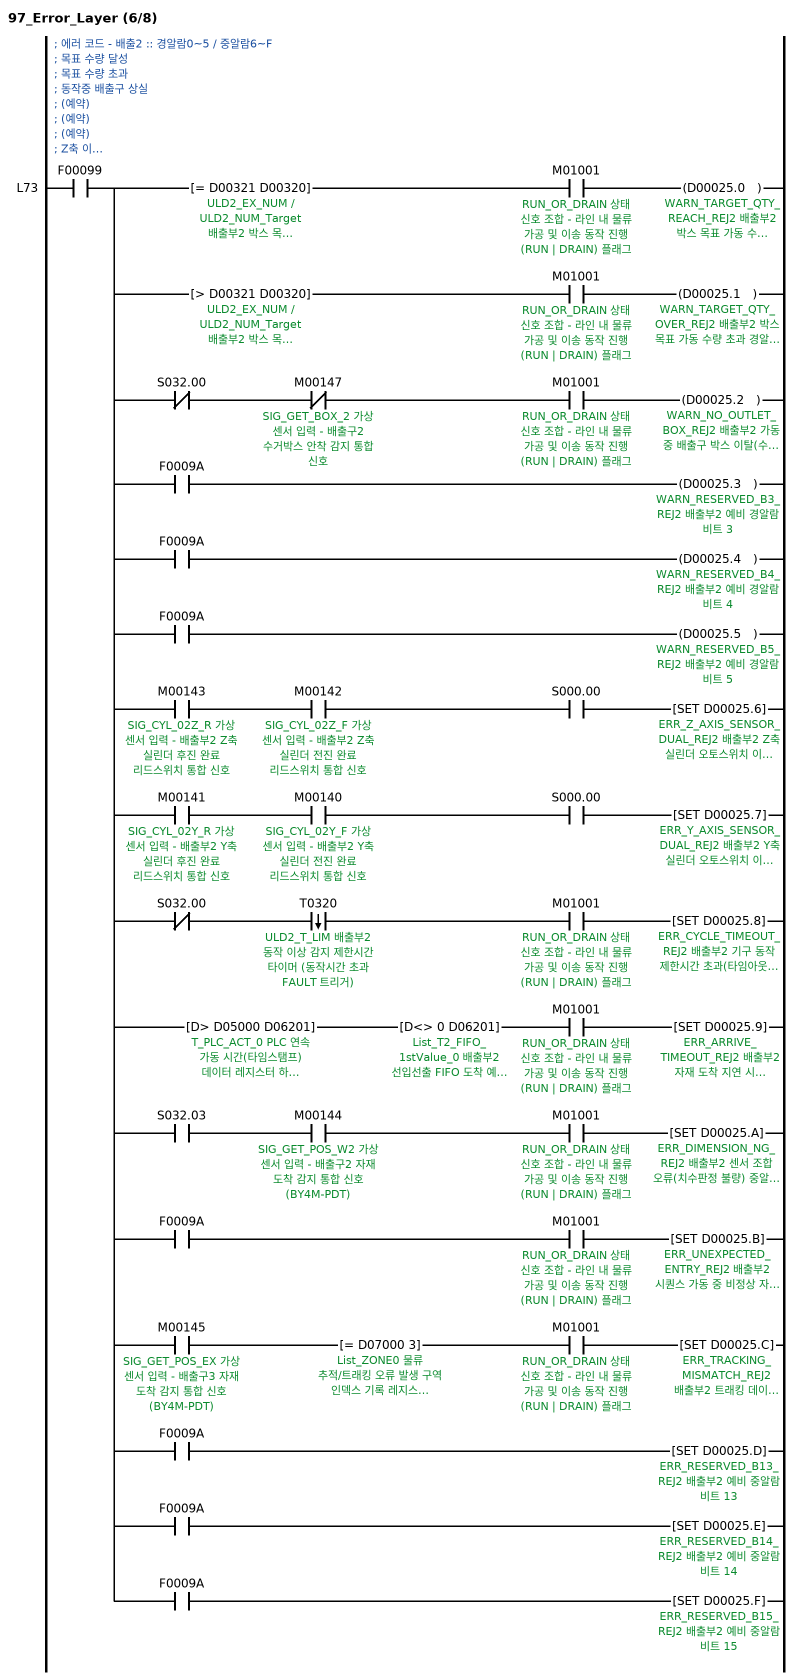
// 에러 코드 - 배출2 :: 경알람0~5 / 중알람6~F
; L73
LOAD      F00099
MPUSH
AND=      D00321 D00320	// ULD2_EX_NUM / ULD2_NUM_Target 배출부2 박스 목표 분류/배출 완료 수량 레지스터
AND       M01001	// RUN_OR_DRAIN 상태 신호 조합 - 라인 내 물류 가공 및 이송 동작 진행 (RUN | DRAIN) 플래그
OUT       D00025.0	// WARN_TARGET_QTY_REACH_REJ2 배출부2 박스 목표 가동 수량 도달(만재 상태) 경알람 비트
MLOAD
AND>      D00321 D00320	// ULD2_EX_NUM / ULD2_NUM_Target 배출부2 박스 목표 분류/배출 완료 수량 레지스터
AND       M01001	// RUN_OR_DRAIN 상태 신호 조합 - 라인 내 물류 가공 및 이송 동작 진행 (RUN | DRAIN) 플래그
OUT       D00025.1	// WARN_TARGET_QTY_OVER_REJ2 배출부2 박스 목표 가동 수량 초과 경알람 비트
MLOAD
AND NOT   S032.00
AND NOT   M00147	// SIG_GET_BOX_2 가상 센서 입력 - 배출구2 수거박스 안착 감지 통합 신호
AND       M01001	// RUN_OR_DRAIN 상태 신호 조합 - 라인 내 물류 가공 및 이송 동작 진행 (RUN | DRAIN) 플래그
OUT       D00025.2	// WARN_NO_OUTLET_BOX_REJ2 배출부2 가동 중 배출구 박스 이탈(수거 상실) 경알람 비트
MLOAD
AND       F0009A
OUT       D00025.3	// WARN_RESERVED_B3_REJ2 배출부2 예비 경알람 비트 3
MLOAD
AND       F0009A
OUT       D00025.4	// WARN_RESERVED_B4_REJ2 배출부2 예비 경알람 비트 4
MLOAD
AND       F0009A
OUT       D00025.5	// WARN_RESERVED_B5_REJ2 배출부2 예비 경알람 비트 5
MLOAD
AND       M00143	// SIG_CYL_02Z_R 가상 센서 입력 - 배출부2 Z축 실린더 후진 완료 리드스위치 통합 신호
AND       M00142	// SIG_CYL_02Z_F 가상 센서 입력 - 배출부2 Z축 실린더 전진 완료 리드스위치 통합 신호
AND       S000.00
SET       D00025.6	// ERR_Z_AXIS_SENSOR_DUAL_REJ2 배출부2 Z축 실린더 오토스위치 이상 (상/하한 센서 동시 ON) 중알람 비트
MLOAD
AND       M00141	// SIG_CYL_02Y_R 가상 센서 입력 - 배출부2 Y축 실린더 후진 완료 리드스위치 통합 신호
AND       M00140	// SIG_CYL_02Y_F 가상 센서 입력 - 배출부2 Y축 실린더 전진 완료 리드스위치 통합 신호
AND       S000.00
SET       D00025.7	// ERR_Y_AXIS_SENSOR_DUAL_REJ2 배출부2 Y축 실린더 오토스위치 이상 (전/후진 센서 동시 ON) 중알람 비트
MLOAD
AND NOT   S032.00
ANDN      T0320	// ULD2_T_LIM 배출부2 동작 이상 감지 제한시간 타이머 (동작시간 초과 FAULT 트리거)
AND       M01001	// RUN_OR_DRAIN 상태 신호 조합 - 라인 내 물류 가공 및 이송 동작 진행 (RUN | DRAIN) 플래그
SET       D00025.8	// ERR_CYCLE_TIMEOUT_REJ2 배출부2 기구 동작 제한시간 초과(타임아웃) 중알람 비트
MLOAD
ANDD>     D05000 D06201	// T_PLC_ACT_0 PLC 연속 가동 시간(타임스탬프) 데이터 레지스터 하위 16비트 (0.1초 해상도) / List_T2_FIFO_1stValue_0 배출부2 선입선출 FIFO 도착 예정 시간 데이터 레지스터 하위 16비트 (32비트 연산)
ANDD<>    0 D06201	// List_T2_FIFO_1stValue_0 배출부2 선입선출 FIFO 도착 예정 시간 데이터 레지스터 하위 16비트 (32비트 연산)
AND       M01001	// RUN_OR_DRAIN 상태 신호 조합 - 라인 내 물류 가공 및 이송 동작 진행 (RUN | DRAIN) 플래그
SET       D00025.9	// ERR_ARRIVE_TIMEOUT_REJ2 배출부2 자재 도착 지연 시간 초과(FIFO 대기시간 초과) 중알람 비트
MLOAD
AND       S032.03
AND       M00144	// SIG_GET_POS_W2 가상 센서 입력 - 배출구2 자재 도착 감지 통합 신호 (BY4M-PDT)
AND       M01001	// RUN_OR_DRAIN 상태 신호 조합 - 라인 내 물류 가공 및 이송 동작 진행 (RUN | DRAIN) 플래그
SET       D00025.A	// ERR_DIMENSION_NG_REJ2 배출부2 센서 조합 오류(치수판정 불량) 중알람 비트
MLOAD
AND       F0009A
AND       M01001	// RUN_OR_DRAIN 상태 신호 조합 - 라인 내 물류 가공 및 이송 동작 진행 (RUN | DRAIN) 플래그
SET       D00025.B	// ERR_UNEXPECTED_ENTRY_REJ2 배출부2 시퀀스 가동 중 비정상 자재 진입 중알람 비트
MLOAD
AND       M00145	// SIG_GET_POS_EX 가상 센서 입력 - 배출구3 자재 도착 감지 통합 신호 (BY4M-PDT)
AND=      D07000 3	// List_ZONE0 물류 추적/트래킹 오류 발생 구역 인덱스 기록 레지스터 (List_ZONE0)
AND       M01001	// RUN_OR_DRAIN 상태 신호 조합 - 라인 내 물류 가공 및 이송 동작 진행 (RUN | DRAIN) 플래그
SET       D00025.C	// ERR_TRACKING_MISMATCH_REJ2 배출부2 트래킹 데이터 불일치(추적 오동작) 중알람 비트
MLOAD
AND       F0009A
SET       D00025.D	// ERR_RESERVED_B13_REJ2 배출부2 예비 중알람 비트 13
MLOAD
AND       F0009A
SET       D00025.E	// ERR_RESERVED_B14_REJ2 배출부2 예비 중알람 비트 14
MPOP
AND       F0009A
SET       D00025.F	// ERR_RESERVED_B15_REJ2 배출부2 예비 중알람 비트 15
// output comment: 목표 수량 달성
// output comment: 목표 수량 초과
// output comment: 동작중 배출구 상실
// output comment: (예약)
// output comment: (예약)
// output comment: (예약)
// output comment: Z축 이상
// output comment: Y축 이상
// output comment: 동작시간 초과
// output comment: 도착시간 초과
// output comment: 치수판정 불량
// output comment: 작동중 투입
// output comment: 추적 불일치
// output comment: (예약)
// output comment: (예약)
// output comment: (예약)

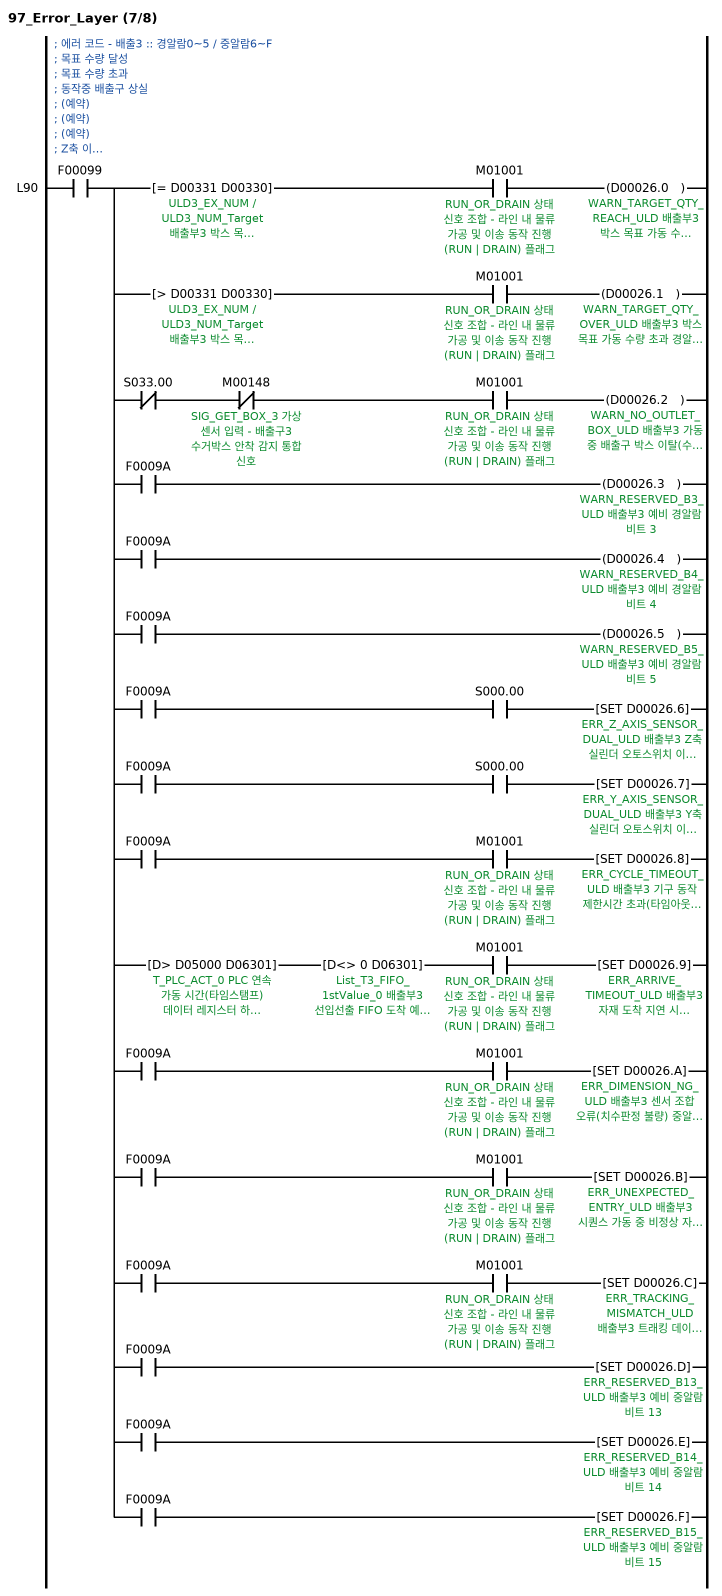
// 에러 코드 - 배출3 :: 경알람0~5 / 중알람6~F
; L90
LOAD      F00099
MPUSH
AND=      D00331 D00330	// ULD3_EX_NUM / ULD3_NUM_Target 배출부3 박스 목표 분류/배출 완료 수량 레지스터
AND       M01001	// RUN_OR_DRAIN 상태 신호 조합 - 라인 내 물류 가공 및 이송 동작 진행 (RUN | DRAIN) 플래그
OUT       D00026.0	// WARN_TARGET_QTY_REACH_ULD 배출부3 박스 목표 가동 수량 도달(만재 상태) 경알람 비트
MLOAD
AND>      D00331 D00330	// ULD3_EX_NUM / ULD3_NUM_Target 배출부3 박스 목표 분류/배출 완료 수량 레지스터
AND       M01001	// RUN_OR_DRAIN 상태 신호 조합 - 라인 내 물류 가공 및 이송 동작 진행 (RUN | DRAIN) 플래그
OUT       D00026.1	// WARN_TARGET_QTY_OVER_ULD 배출부3 박스 목표 가동 수량 초과 경알람 비트
MLOAD
AND NOT   S033.00
AND NOT   M00148	// SIG_GET_BOX_3 가상 센서 입력 - 배출구3 수거박스 안착 감지 통합 신호
AND       M01001	// RUN_OR_DRAIN 상태 신호 조합 - 라인 내 물류 가공 및 이송 동작 진행 (RUN | DRAIN) 플래그
OUT       D00026.2	// WARN_NO_OUTLET_BOX_ULD 배출부3 가동 중 배출구 박스 이탈(수거 상실) 경알람 비트
MLOAD
AND       F0009A
OUT       D00026.3	// WARN_RESERVED_B3_ULD 배출부3 예비 경알람 비트 3
MLOAD
AND       F0009A
OUT       D00026.4	// WARN_RESERVED_B4_ULD 배출부3 예비 경알람 비트 4
MLOAD
AND       F0009A
OUT       D00026.5	// WARN_RESERVED_B5_ULD 배출부3 예비 경알람 비트 5
MLOAD
AND       F0009A
AND       S000.00
SET       D00026.6	// ERR_Z_AXIS_SENSOR_DUAL_ULD 배출부3 Z축 실린더 오토스위치 이상 (상/하한 센서 동시 ON) 중알람 비트
MLOAD
AND       F0009A
AND       S000.00
SET       D00026.7	// ERR_Y_AXIS_SENSOR_DUAL_ULD 배출부3 Y축 실린더 오토스위치 이상 (전/후진 센서 동시 ON) 중알람 비트
MLOAD
AND       F0009A
AND       M01001	// RUN_OR_DRAIN 상태 신호 조합 - 라인 내 물류 가공 및 이송 동작 진행 (RUN | DRAIN) 플래그
SET       D00026.8	// ERR_CYCLE_TIMEOUT_ULD 배출부3 기구 동작 제한시간 초과(타임아웃) 중알람 비트
MLOAD
ANDD>     D05000 D06301	// T_PLC_ACT_0 PLC 연속 가동 시간(타임스탬프) 데이터 레지스터 하위 16비트 (0.1초 해상도) / List_T3_FIFO_1stValue_0 배출부3 선입선출 FIFO 도착 예정 시간 데이터 레지스터 하위 16비트 (32비트 연산)
ANDD<>    0 D06301	// List_T3_FIFO_1stValue_0 배출부3 선입선출 FIFO 도착 예정 시간 데이터 레지스터 하위 16비트 (32비트 연산)
AND       M01001	// RUN_OR_DRAIN 상태 신호 조합 - 라인 내 물류 가공 및 이송 동작 진행 (RUN | DRAIN) 플래그
SET       D00026.9	// ERR_ARRIVE_TIMEOUT_ULD 배출부3 자재 도착 지연 시간 초과(FIFO 대기시간 초과) 중알람 비트
MLOAD
AND       F0009A
AND       M01001	// RUN_OR_DRAIN 상태 신호 조합 - 라인 내 물류 가공 및 이송 동작 진행 (RUN | DRAIN) 플래그
SET       D00026.A	// ERR_DIMENSION_NG_ULD 배출부3 센서 조합 오류(치수판정 불량) 중알람 비트
MLOAD
AND       F0009A
AND       M01001	// RUN_OR_DRAIN 상태 신호 조합 - 라인 내 물류 가공 및 이송 동작 진행 (RUN | DRAIN) 플래그
SET       D00026.B	// ERR_UNEXPECTED_ENTRY_ULD 배출부3 시퀀스 가동 중 비정상 자재 진입 중알람 비트
MLOAD
AND       F0009A
AND       M01001	// RUN_OR_DRAIN 상태 신호 조합 - 라인 내 물류 가공 및 이송 동작 진행 (RUN | DRAIN) 플래그
SET       D00026.C	// ERR_TRACKING_MISMATCH_ULD 배출부3 트래킹 데이터 불일치(추적 오동작) 중알람 비트
MLOAD
AND       F0009A
SET       D00026.D	// ERR_RESERVED_B13_ULD 배출부3 예비 중알람 비트 13
MLOAD
AND       F0009A
SET       D00026.E	// ERR_RESERVED_B14_ULD 배출부3 예비 중알람 비트 14
MPOP
AND       F0009A
SET       D00026.F	// ERR_RESERVED_B15_ULD 배출부3 예비 중알람 비트 15
// output comment: 목표 수량 달성
// output comment: 목표 수량 초과
// output comment: 동작중 배출구 상실
// output comment: (예약)
// output comment: (예약)
// output comment: (예약)
// output comment: Z축 이상
// output comment: Y축 이상
// output comment: 동작시간 초과
// output comment: 도착시간 초과
// output comment: 치수판정 불량
// output comment: 작동중 투입
// output comment: 추적 불일치
// output comment: (예약)
// output comment: (예약)
// output comment: (예약)

